// TIA Portal V21 program export: 0 tag tables, 0 data types, 1 data blocks, 40 code blocks (in call order from the OBs), 24 instance data blocks

DATA_BLOCK "Global_Limits_Interlocks"   // DB58
{ S7_Optimized_Access := 'TRUE' }
// stored: MemoryReserve 100
   VAR
      ExternalLevel_Interlock : Real := 2900.0;
      InternalLevel_Interlock : Real := 2700.0;
   END_VAR
BEGIN
END_DATA_BLOCK

ORGANIZATION_BLOCK "Main_1"   // OB1, LAD, ProgramCycle
TITLE = "Main Program Sweep (Cycle)"
{ S7_Optimized_Access := 'TRUE' }
// stored: SetENOAutomatically false
   VAR_INPUT
      Initial_Call : Bool;   // Initial call of this OB
      Remanence : Bool;   // =True, if remanent data are available
   END_VAR
BEGIN
END_ORGANIZATION_BLOCK

ORGANIZATION_BLOCK "Cyclic interrupt"   // OB30, FBD, CyclicInterrupt
{ S7_Optimized_Access := 'TRUE' }
// stored: SetENOAutomatically false
   VAR_INPUT
      Initial_Call : Bool;   // Initial call of this OB
      Event_Count : Int;   // Events discarded
   END_VAR
BEGIN

REGION Network 1: Service
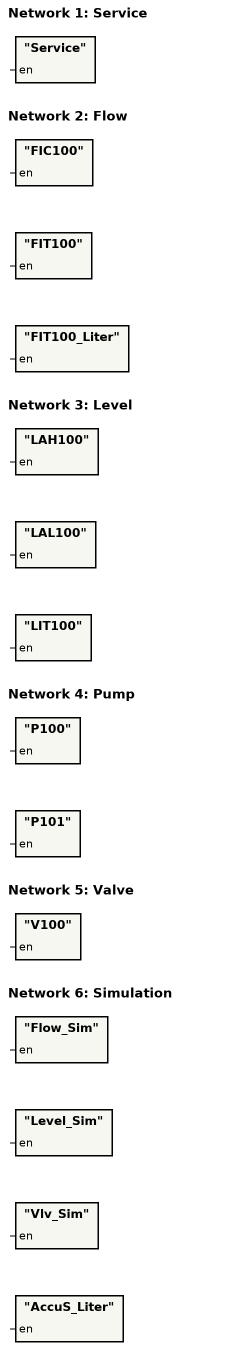
   "Service"();
END_REGION

REGION Network 2: Flow
   "FIC100"();
   "FIT100"();
   "FIT100_Liter"();
END_REGION

REGION Network 3: Level
   "LAH100"();
   "LAL100"();
   "LIT100"();
END_REGION

REGION Network 4: Pump
   "P100"();
   "P101"();
END_REGION

REGION Network 5: Valve
   "V100"();
END_REGION

REGION Network 6: Simulation
   "Flow_Sim"();
   "Level_Sim"();
   "Vlv_Sim"();
   "AccuS_Liter"();
END_REGION
END_ORGANIZATION_BLOCK

FUNCTION "Service" : Void   // FC11, FBD
TITLE = Service
{ S7_Optimized_Access := 'TRUE' }
AUTHOR : Siemens AG
FAMILY : ServiceControl
VERSION : 1.0
// stored: SetENOAutomatically false
   VAR_TEMP
      ProcedureDone : Bool;
      UnholdingDone : Bool;
      StartingState : Bool;
      CompletingState : Bool;
      PausingState : Bool;
      HoldingState : Bool;
      AbortingState : Bool;
      StoppingState : Bool;
      State : "Service_States";
   END_VAR
   VAR_TEMP   // added for the SCL form of the ladder/FBD networks
      _w1 : Bool;
      _w2 : Bool;
      _w3 : Bool;
      _w4 : Bool;
   END_VAR
BEGIN

REGION Network 1: Parameters and values
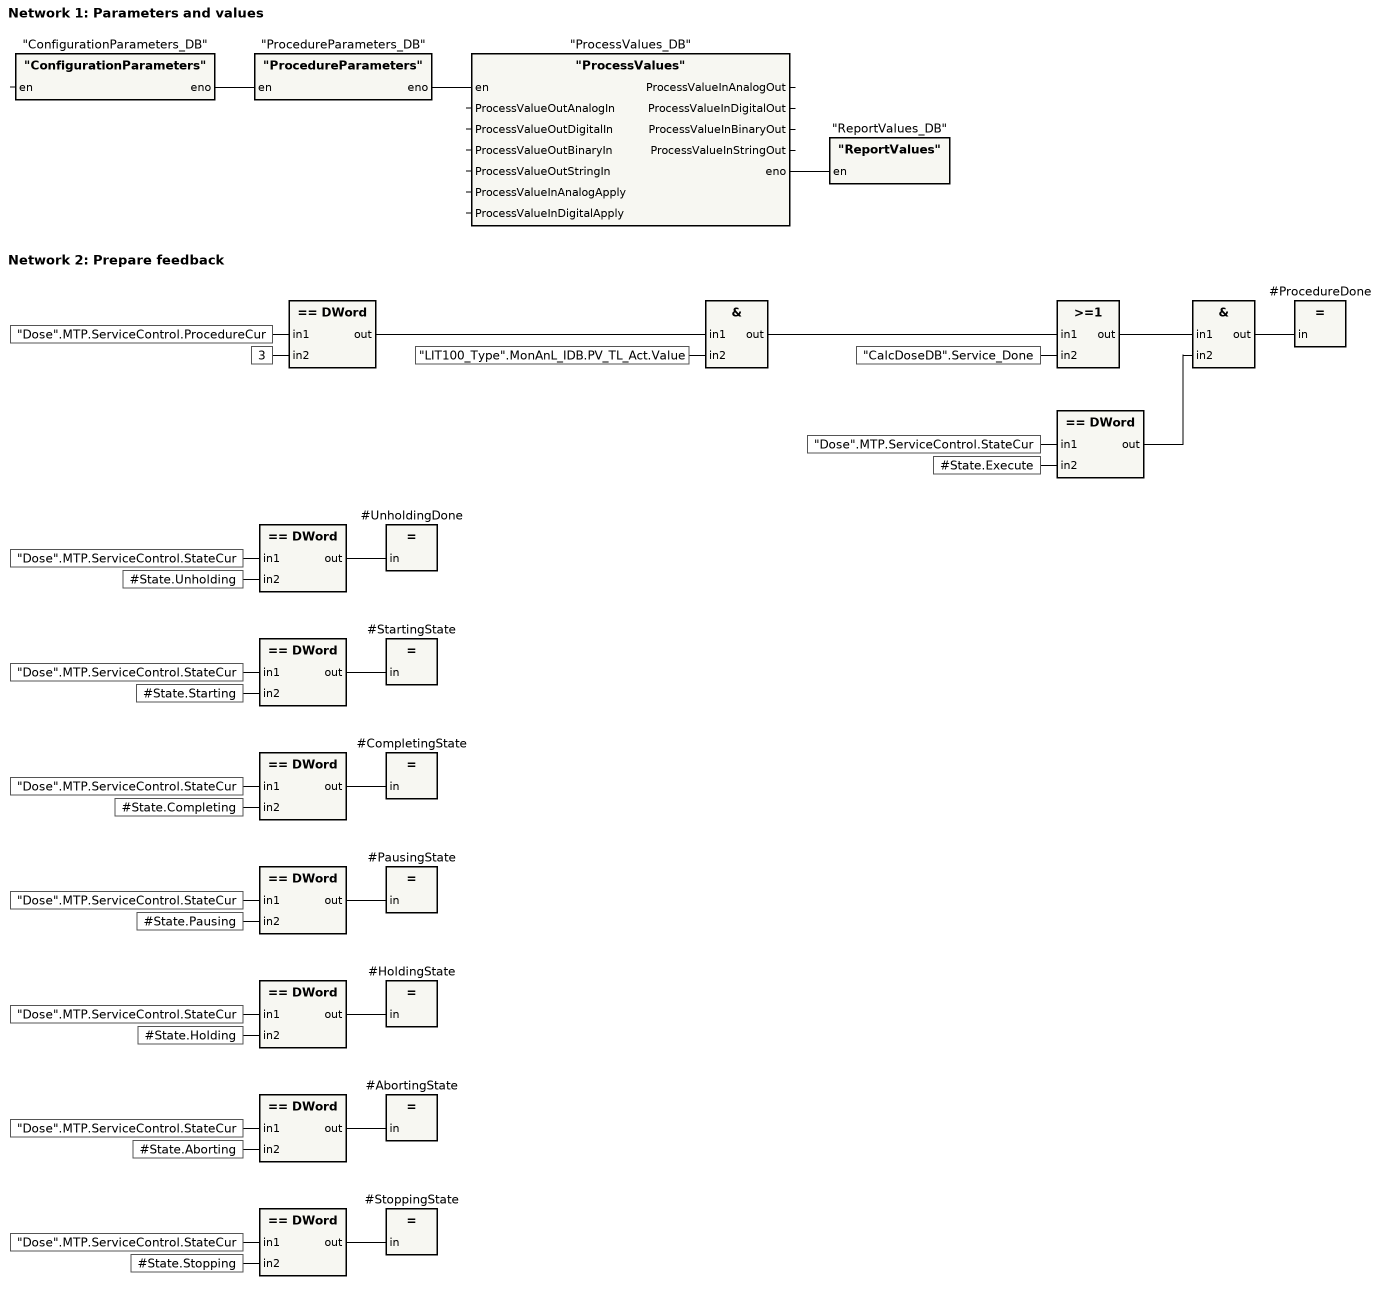
   "ConfigurationParameters_DB"(ENO => #_w1);   // "ConfigurationParameters"
   "ProcedureParameters_DB"(EN := #_w1, ENO => #_w2);   // "ProcedureParameters"
   "ProcessValues_DB"(EN := #_w2, ENO => #_w3);   // "ProcessValues"
   IF #_w3 THEN
       "ReportValues_DB"();   // "ReportValues"
   END_IF;
END_REGION

REGION Network 2: Prepare feedback
   #ProcedureDone := ((("Dose".MTP.ServiceControl.ProcedureCur = 3) AND "LIT100_Type".MonAnL_IDB.PV_TL_Act.Value) OR "CalcDoseDB".Service_Done) AND ("Dose".MTP.ServiceControl.StateCur = #State.Execute);
   #UnholdingDone := "Dose".MTP.ServiceControl.StateCur = #State.Unholding;
   #StartingState := "Dose".MTP.ServiceControl.StateCur = #State.Starting;
   #CompletingState := "Dose".MTP.ServiceControl.StateCur = #State.Completing;
   #PausingState := "Dose".MTP.ServiceControl.StateCur = #State.Pausing;
   #HoldingState := "Dose".MTP.ServiceControl.StateCur = #State.Holding;
   #AbortingState := "Dose".MTP.ServiceControl.StateCur = #State.Aborting;
   #StoppingState := "Dose".MTP.ServiceControl.StateCur = #State.Stopping;
END_REGION

REGION Network 3: Cm P100 feedback
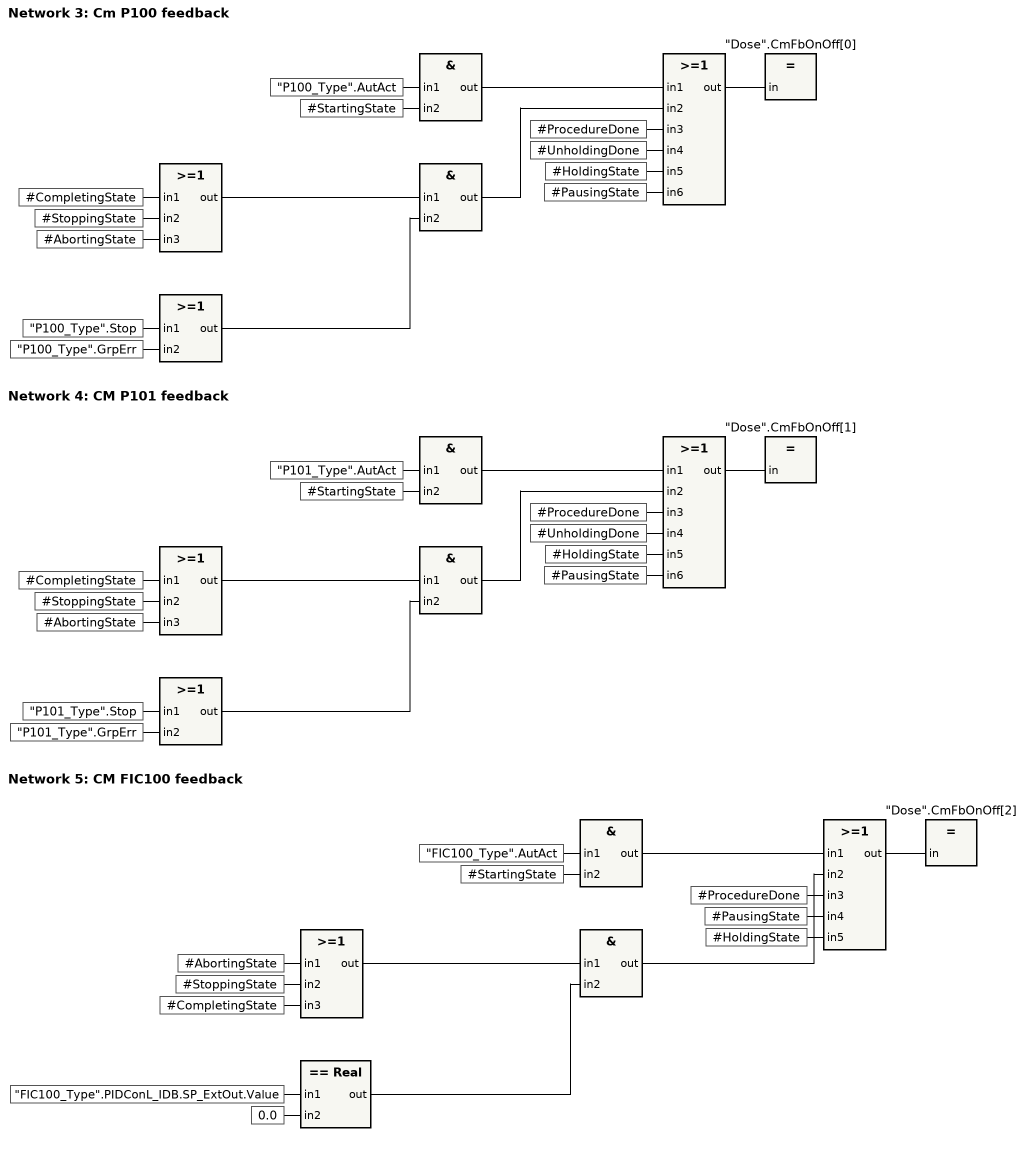
   "Dose".CmFbOnOff[0] := ("P100_Type".AutAct AND #StartingState) OR ((#CompletingState OR #StoppingState OR #AbortingState) AND ("P100_Type".Stop OR "P100_Type".GrpErr)) OR #ProcedureDone OR #UnholdingDone OR #HoldingState OR #PausingState;
END_REGION

REGION Network 4: CM P101 feedback
   "Dose".CmFbOnOff[1] := ("P101_Type".AutAct AND #StartingState) OR ((#CompletingState OR #StoppingState OR #AbortingState) AND ("P101_Type".Stop OR "P101_Type".GrpErr)) OR #ProcedureDone OR #UnholdingDone OR #HoldingState OR #PausingState;
END_REGION

REGION Network 5: CM FIC100 feedback
   "Dose".CmFbOnOff[2] := ("FIC100_Type".AutAct AND #StartingState) OR ((#AbortingState OR #StoppingState OR #CompletingState) AND ("FIC100_Type".PIDConL_IDB.SP_ExtOut.Value = 0.0)) OR #ProcedureDone OR #PausingState OR #HoldingState;
END_REGION

REGION Network 6: CM V100 feedback
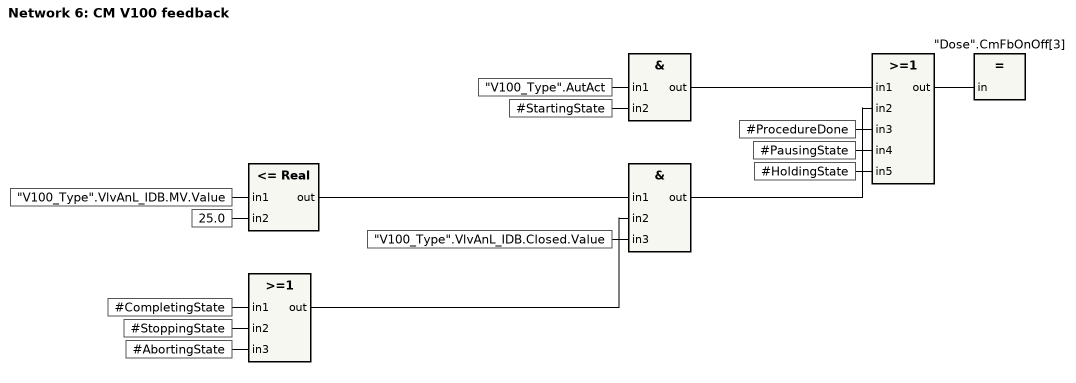
   "Dose".CmFbOnOff[3] := ("V100_Type".AutAct AND #StartingState) OR (("V100_Type".VlvAnL_IDB.MV.Value <= 25.0) AND (#CompletingState OR #StoppingState OR #AbortingState) AND "V100_Type".VlvAnL_IDB.Closed.Value) OR #ProcedureDone OR #PausingState OR #HoldingState;
END_REGION

REGION Network 7: Service
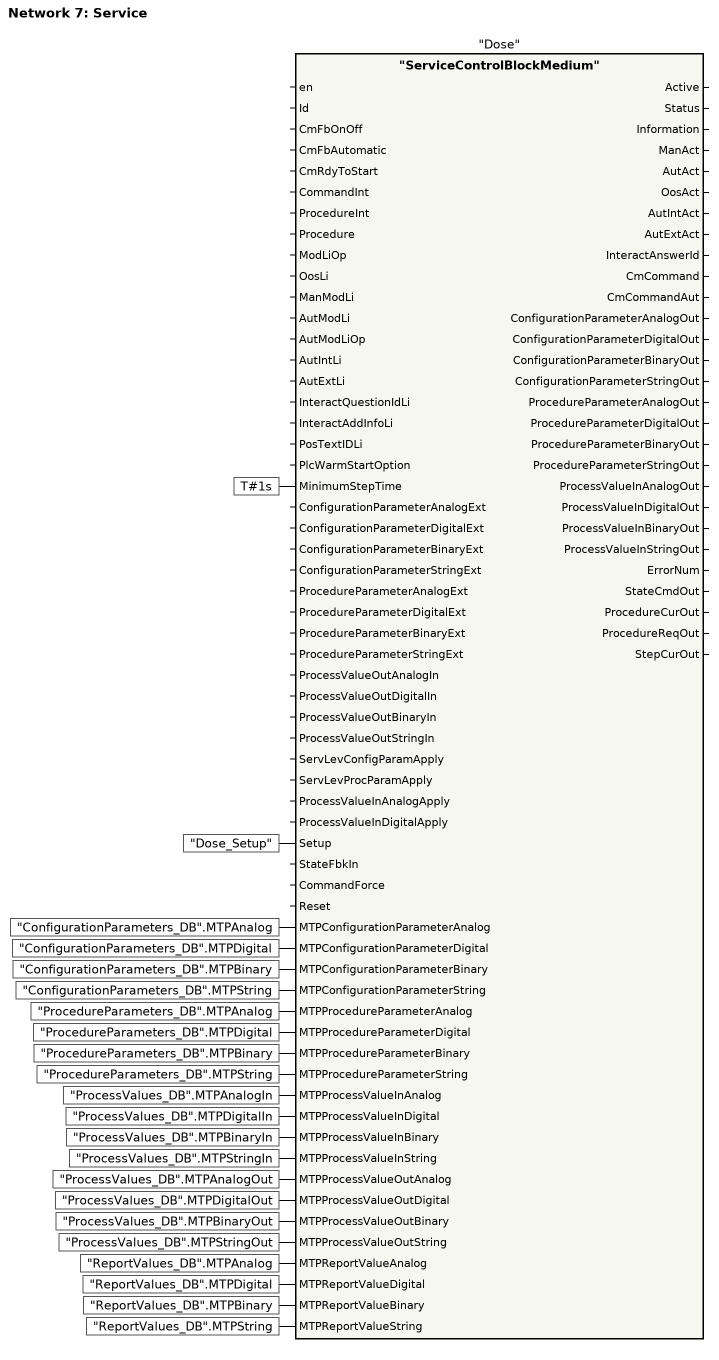
   "Dose"(MinimumStepTime := T#1s,   // "ServiceControlBlockMedium"
          Setup := "Dose_Setup",
          MTPConfigurationParameterAnalog := "ConfigurationParameters_DB".MTPAnalog,
          MTPConfigurationParameterDigital := "ConfigurationParameters_DB".MTPDigital,
          MTPConfigurationParameterBinary := "ConfigurationParameters_DB".MTPBinary,
          MTPConfigurationParameterString := "ConfigurationParameters_DB".MTPString,
          MTPProcedureParameterAnalog := "ProcedureParameters_DB".MTPAnalog,
          MTPProcedureParameterDigital := "ProcedureParameters_DB".MTPDigital,
          MTPProcedureParameterBinary := "ProcedureParameters_DB".MTPBinary,
          MTPProcedureParameterString := "ProcedureParameters_DB".MTPString,
          MTPProcessValueInAnalog := "ProcessValues_DB".MTPAnalogIn,
          MTPProcessValueInDigital := "ProcessValues_DB".MTPDigitalIn,
          MTPProcessValueInBinary := "ProcessValues_DB".MTPBinaryIn,
          MTPProcessValueInString := "ProcessValues_DB".MTPStringIn,
          MTPProcessValueOutAnalog := "ProcessValues_DB".MTPAnalogOut,
          MTPProcessValueOutDigital := "ProcessValues_DB".MTPDigitalOut,
          MTPProcessValueOutBinary := "ProcessValues_DB".MTPBinaryOut,
          MTPProcessValueOutString := "ProcessValues_DB".MTPStringOut,
          MTPReportValueAnalog := "ReportValues_DB".MTPAnalog,
          MTPReportValueDigital := "ReportValues_DB".MTPDigital,
          MTPReportValueBinary := "ReportValues_DB".MTPBinary,
          MTPReportValueString := "ReportValues_DB".MTPString);
END_REGION

REGION Network 8: Service HMI
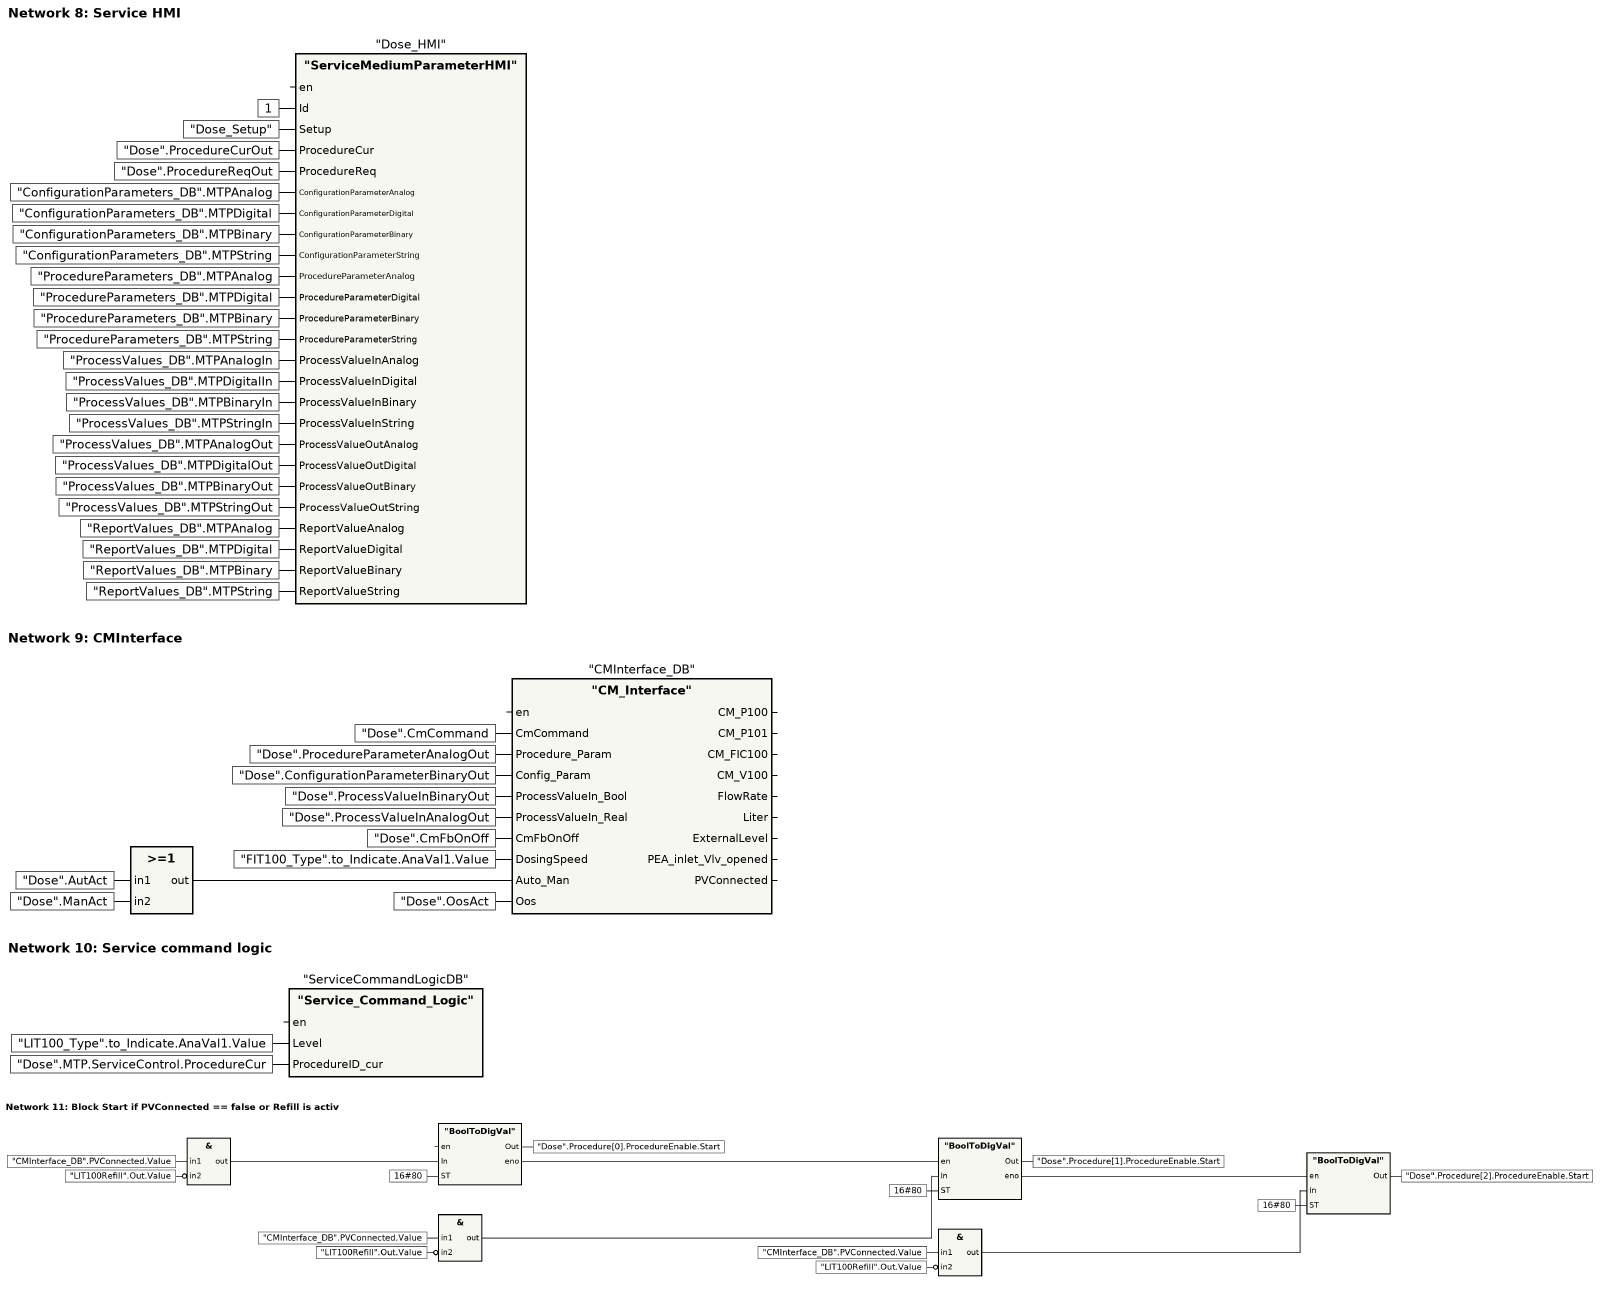
   "Dose_HMI"(Id := 1,   // "ServiceMediumParameterHMI"
              Setup := "Dose_Setup",
              ProcedureCur := "Dose".ProcedureCurOut,
              ProcedureReq := "Dose".ProcedureReqOut,
              ConfigurationParameterAnalog := "ConfigurationParameters_DB".MTPAnalog,
              ConfigurationParameterDigital := "ConfigurationParameters_DB".MTPDigital,
              ConfigurationParameterBinary := "ConfigurationParameters_DB".MTPBinary,
              ConfigurationParameterString := "ConfigurationParameters_DB".MTPString,
              ProcedureParameterAnalog := "ProcedureParameters_DB".MTPAnalog,
              ProcedureParameterDigital := "ProcedureParameters_DB".MTPDigital,
              ProcedureParameterBinary := "ProcedureParameters_DB".MTPBinary,
              ProcedureParameterString := "ProcedureParameters_DB".MTPString,
              ProcessValueInAnalog := "ProcessValues_DB".MTPAnalogIn,
              ProcessValueInDigital := "ProcessValues_DB".MTPDigitalIn,
              ProcessValueInBinary := "ProcessValues_DB".MTPBinaryIn,
              ProcessValueInString := "ProcessValues_DB".MTPStringIn,
              ProcessValueOutAnalog := "ProcessValues_DB".MTPAnalogOut,
              ProcessValueOutDigital := "ProcessValues_DB".MTPDigitalOut,
              ProcessValueOutBinary := "ProcessValues_DB".MTPBinaryOut,
              ProcessValueOutString := "ProcessValues_DB".MTPStringOut,
              ReportValueAnalog := "ReportValues_DB".MTPAnalog,
              ReportValueDigital := "ReportValues_DB".MTPDigital,
              ReportValueBinary := "ReportValues_DB".MTPBinary,
              ReportValueString := "ReportValues_DB".MTPString);
END_REGION

REGION Network 9: CMInterface
   "CMInterface_DB"(CmCommand := "Dose".CmCommand,   // "CM_Interface"
                    Procedure_Param := "Dose".ProcedureParameterAnalogOut,
                    Config_Param := "Dose".ConfigurationParameterBinaryOut,
                    ProcessValueIn_Bool := "Dose".ProcessValueInBinaryOut,
                    ProcessValueIn_Real := "Dose".ProcessValueInAnalogOut,
                    CmFbOnOff := "Dose".CmFbOnOff,
                    DosingSpeed := "FIT100_Type".to_Indicate.AnaVal1.Value,
                    Auto_Man := "Dose".AutAct OR "Dose".ManAct,
                    Oos := "Dose".OosAct);
END_REGION

REGION Network 10: Service command logic
   "ServiceCommandLogicDB"(Level := "LIT100_Type".to_Indicate.AnaVal1.Value,   // "Service_Command_Logic"
                           ProcedureID_cur := "Dose".MTP.ServiceControl.ProcedureCur);
END_REGION

REGION Network 11: Block Start if PVConnected == false or Refill is activ
   "BoolToDigVal"(In := "CMInterface_DB".PVConnected.Value AND NOT "LIT100Refill".Out.Value,
                  ST := 16#80,
                  Out => "Dose".Procedure[0].ProcedureEnable.Start,
                  ENO => #_w1);
   "BoolToDigVal"(EN := #_w1,
                  In := "CMInterface_DB".PVConnected.Value AND NOT "LIT100Refill".Out.Value,
                  ST := 16#80,
                  Out => "Dose".Procedure[1].ProcedureEnable.Start,
                  ENO => #_w2);
   IF #_w2 THEN
       "BoolToDigVal"(In := "CMInterface_DB".PVConnected.Value AND NOT "LIT100Refill".Out.Value,
                      ST := 16#80,
                      Out => "Dose".Procedure[2].ProcedureEnable.Start);
   END_IF;
END_REGION

REGION Network 12: Block Resume and Unholding if refill is activ
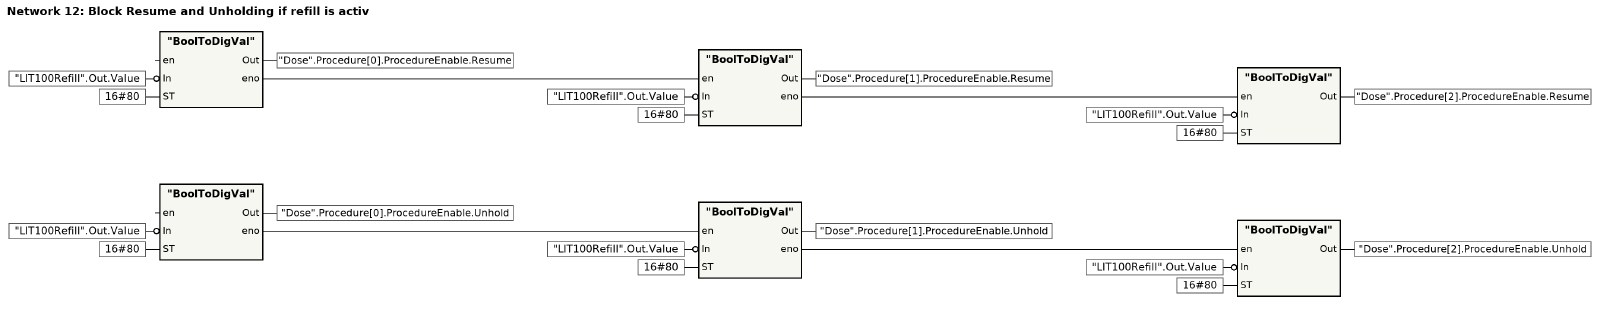
   "BoolToDigVal"(In := NOT "LIT100Refill".Out.Value,
                  ST := 16#80,
                  Out => "Dose".Procedure[0].ProcedureEnable.Resume,
                  ENO => #_w1);
   "BoolToDigVal"(EN := #_w1,
                  In := NOT "LIT100Refill".Out.Value,
                  ST := 16#80,
                  Out => "Dose".Procedure[1].ProcedureEnable.Resume,
                  ENO => #_w2);
   IF #_w2 THEN
       "BoolToDigVal"(In := NOT "LIT100Refill".Out.Value,
                      ST := 16#80,
                      Out => "Dose".Procedure[2].ProcedureEnable.Resume);
   END_IF;
   "BoolToDigVal"(In := NOT "LIT100Refill".Out.Value,
                  ST := 16#80,
                  Out => "Dose".Procedure[0].ProcedureEnable.Unhold,
                  ENO => #_w3);
   "BoolToDigVal"(EN := #_w3,
                  In := NOT "LIT100Refill".Out.Value,
                  ST := 16#80,
                  Out => "Dose".Procedure[1].ProcedureEnable.Unhold,
                  ENO => #_w4);
   IF #_w4 THEN
       "BoolToDigVal"(In := NOT "LIT100Refill".Out.Value,
                      ST := 16#80,
                      Out => "Dose".Procedure[2].ProcedureEnable.Unhold);
   END_IF;
END_REGION

REGION Network 13: Position Text
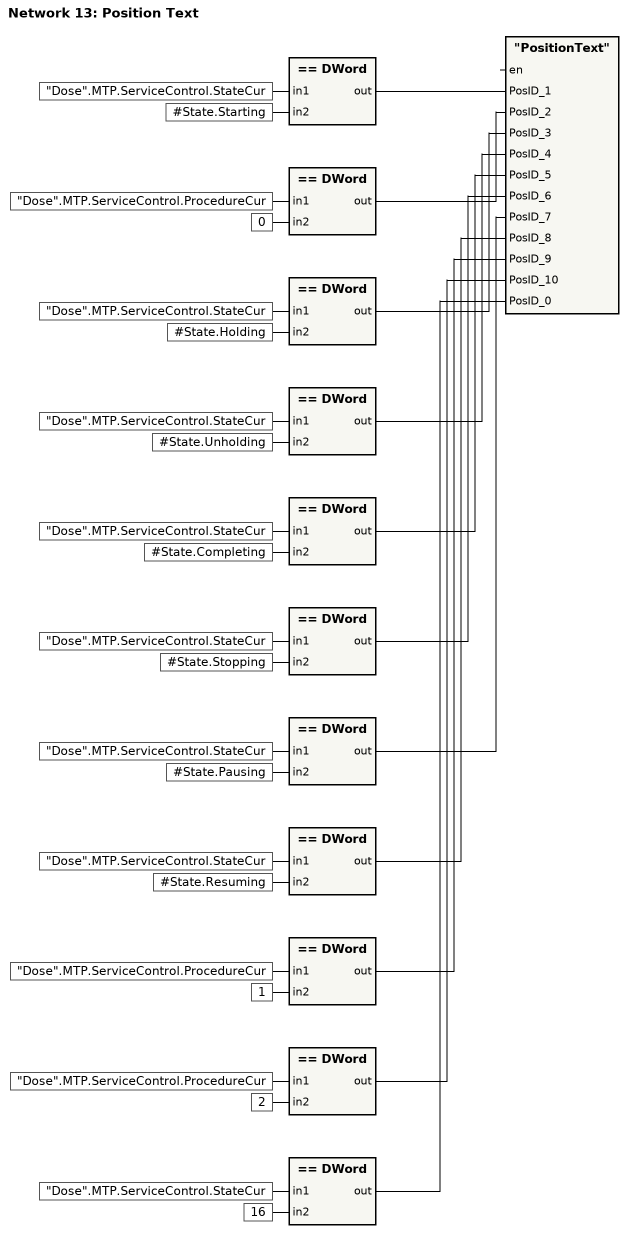
   "PositionText"(PosID_1 := "Dose".MTP.ServiceControl.StateCur = #State.Starting,
                  PosID_2 := "Dose".MTP.ServiceControl.ProcedureCur = 0,
                  PosID_3 := "Dose".MTP.ServiceControl.StateCur = #State.Holding,
                  PosID_4 := "Dose".MTP.ServiceControl.StateCur = #State.Unholding,
                  PosID_5 := "Dose".MTP.ServiceControl.StateCur = #State.Completing,
                  PosID_6 := "Dose".MTP.ServiceControl.StateCur = #State.Stopping,
                  PosID_7 := "Dose".MTP.ServiceControl.StateCur = #State.Pausing,
                  PosID_8 := "Dose".MTP.ServiceControl.StateCur = #State.Resuming,
                  PosID_9 := "Dose".MTP.ServiceControl.ProcedureCur = 1,
                  PosID_10 := "Dose".MTP.ServiceControl.ProcedureCur = 2,
                  PosID_0 := "Dose".MTP.ServiceControl.StateCur = 16);
END_REGION

REGION Network 14: Report values
END_REGION
END_FUNCTION

FUNCTION_BLOCK "ConfigurationParameters"   // FB1710, SCL
TITLE = ConfigurationParameters
{ S7_Optimized_Access := 'TRUE' }
AUTHOR : Siemens AG
FAMILY : ServiceControl
VERSION : 1.0
// Providing of the MTP-Interface and the number of parameters of each configuration parameter type
// stored: MemoryReserve 100, SetENOAutomatically false
   VAR
      MTPAnalog { S7_SetPoint := 'True'} : Array[0..#NUMBER_PARAMETERS_ANALOG] of "UDT_MTP_AnaServParam";
      MTPDigital { S7_SetPoint := 'True'} : Array[0..#NUMBER_PARAMETERS_DIGITAL] of "UDT_MTP_DIntServParam";
      MTPBinary { S7_SetPoint := 'True'} : Array[0..#NUMBER_PARAMETERS_BINARY] of "UDT_MTP_BinServParam";
      MTPString { S7_SetPoint := 'True'} : Array[0..#NUMBER_PARAMETERS_STRING] of "UDT_MTP_StringServParam";
   END_VAR
   VAR CONSTANT
      NUMBER_PARAMETERS_ANALOG : Int := 0;
      NUMBER_PARAMETERS_DIGITAL : Int := 0;
      NUMBER_PARAMETERS_BINARY : Int := 1;
      NUMBER_PARAMETERS_STRING : Int := 0;
   END_VAR
BEGIN
   REGION Block Info Header
     //===============================================================================
     // Siemens AG / (c)Copyright 2021
     //-------------------------------------------------------------------------------
     // Title:            ConfigurationParameters
     // Comment/Function: Providing of the MTP-Interface and the number of parameters of each configuration parameter type
     // Library/Family:   ServiceControl
     // Author:           Siemens AG
     // Tested with:      S7-PLCSIM Advanced 4.0
     // Engineering:      TIA Portal V17
     // Restrictions:     MTP
     // Requirements:     PLC (S7-1200 / S7-1500)
     //-------------------------------------------------------------------------------
     // Change log table:
     // Version  | Date       | Expert in charge        | Changes applied
     //----------|------------|-------------------------|-----------------------------
     // 01.00.00 | 02.09.2021 | Michael Schlosser       | First released version
     // 01.00.01 | 07.09.2021 | Michael Schlosser       | Change: Interface of FB28 ConfigurationParameterAnalog
     // 01.00.02 | 08.09.2021 | Michael Schlosser       | Change: Interface of FB18, FB33, FB24
     // 01.00.03 | 09.09.2021 | Michael Schlosser       | Change: For-loops only until #NUMBER_PARAMETERS_YXZ - 1
     // 01.00.04 | 15.09.2021 | Michael Schlosser       | Change: ApplyEn default values = true (e.g. parLevAnalogApplyEn[0])
     // 01.00.05 | 16.09.2021 | Michael Schlosser       | Change: ApplyEn & ApplyInt as part of UDT_Service_ParameterApply (e.g. #ParLevAnalogApply[0].En)
     // 01.00.06 | 18.10.2021 | Michael Schlosser       | change: call of FBs for parameters now in ServiceControlBlock-FBs to allow several services per PLC
     //===============================================================================
   END_REGION Block Info Header

   REGION Description
     // ConfigurationParameters provides the MTP-Interface and the number of parameters of each configuration parameter type
   END_REGION Description
END_FUNCTION_BLOCK

FUNCTION_BLOCK "ProcedureParameters"   // FB1715, SCL
TITLE = ProcedureParameters
{ S7_Optimized_Access := 'TRUE' }
AUTHOR : Siemens AG
FAMILY : ServiceControl
VERSION : 1.0
// Providing of the MTP-Interface and the number of parameters of each procedure parameter type
// stored: MemoryReserve 100, SetENOAutomatically false
   VAR
      MTPAnalog { S7_SetPoint := 'True'} : Array[0..#NUMBER_PARAMETERS_ANALOG] of "UDT_MTP_AnaServParam";
      MTPDigital { S7_SetPoint := 'True'} : Array[0..#NUMBER_PARAMETERS_DIGITAL] of "UDT_MTP_DIntServParam";
      MTPBinary { S7_SetPoint := 'True'} : Array[0..#NUMBER_PARAMETERS_BINARY] of "UDT_MTP_BinServParam";
      MTPString { S7_SetPoint := 'True'} : Array[0..#NUMBER_PARAMETERS_STRING] of "UDT_MTP_StringServParam";
   END_VAR
   VAR CONSTANT
      NUMBER_PARAMETERS_ANALOG : Int := 2;
      NUMBER_PARAMETERS_DIGITAL : Int := 0;
      NUMBER_PARAMETERS_BINARY : Int := 0;
      NUMBER_PARAMETERS_STRING : Int := 0;
   END_VAR
BEGIN
   REGION Block Info Header
     //===============================================================================
     // Siemens AG / (c)Copyright 2021
     //-------------------------------------------------------------------------------
     // Title:            ProcedureParameters
     // Comment/Function: Providing of the MTP-Interface and the number of parameters of each procedure parameter type
     // Library/Family:   ServiceControl
     // Author:           Siemens AG
     // Tested with:      S7-PLCSIM Advanced 4.0
     // Engineering:      TIA Portal V17
     // Restrictions:     MTP
     // Requirements:     PLC (S7-1200 / S7-1500)
     //-------------------------------------------------------------------------------
     // Change log table:
     // Version  | Date       | Expert in charge        | Changes applied
     //----------|------------|-------------------------|-----------------------------
     // 01.00.00 | 02.09.2021 | Michael Schlosser       | First released version
     // 01.00.01 | 13.09.2021 | Michael Schlosser       | Change: Interface of FB29
     // 01.00.02 | 15.09.2021 | Michael Schlosser       | Change: Interface of FB13, FB19, FB23
     // 01.00.03 | 15.09.2021 | Michael Schlosser       | Change: ApplyEn default values = true (e.g. parLevAnalogApplyEn[0])
     // 01.00.04 | 16.09.2021 | Michael Schlosser       | Change: ApplyEn & ApplyInt as part of UDT_Service_ParameterApply (e.g. #ParLevAnalogApply[0].En)
     // 01.00.05 | 18.10.2021 | Michael Schlosser       | change: call of FBs for parameters now in ServiceControlBlock-FBs to allow several services per PLC
     //===============================================================================
   END_REGION Block Info Header

   REGION Description
     // ProcedureParameters provides the MTP-Interface and the number of parameters of each procedure parameter type
   END_REGION Description
END_FUNCTION_BLOCK

FUNCTION_BLOCK "ProcessValues"   // FB1720, SCL
TITLE = ProcessValues
{ S7_Optimized_Access := 'TRUE' }
AUTHOR : Siemens AG
FAMILY : ServiceControl
VERSION : 1.0
// Handling of ProcessValues
// stored: MemoryReserve 100, SetENOAutomatically false
   VAR_INPUT
      ProcessValueOutAnalogIn { ExternalAccessible := 'False'; ExternalVisible := 'False'; ExternalWritable := 'False'} : Array[0..#NUMBER_PARAMETERS_OUT_ANALOG_NOT_MAPPED] of "UDT_MTP_AnaProcessValueOut";
      ProcessValueOutDigitalIn { ExternalAccessible := 'False'; ExternalVisible := 'False'; ExternalWritable := 'False'} : Array[0..#NUMBER_PARAMETERS_OUT_DIGITAL_NOT_MAPPED] of "UDT_MTP_DIntProcessValueOut";
      ProcessValueOutBinaryIn { ExternalAccessible := 'False'; ExternalVisible := 'False'; ExternalWritable := 'False'} : Array[0..#NUMBER_PARAMETERS_OUT_BINARY_NOT_MAPPED] of "UDT_MTP_BinProcessValueOut";
      ProcessValueOutStringIn { ExternalAccessible := 'False'; ExternalVisible := 'False'; ExternalWritable := 'False'} : Array[0..#NUMBER_PARAMETERS_OUT_STRING_NOT_MAPPED] of "UDT_MTP_StringProcessValueOut";
      ProcessValueInAnalogApply { ExternalAccessible := 'False'; ExternalVisible := 'False'; ExternalWritable := 'False'} : Array[0..#NUMBER_PARAMETERS_IN_ANALOG_NOT_MAPPED] of "UDT_Service_ProcessValueInApply";
      ProcessValueInDigitalApply { ExternalAccessible := 'False'; ExternalVisible := 'False'; ExternalWritable := 'False'} : Array[0..#NUMBER_PARAMETERS_IN_DIGITAL_NOT_MAPPED] of "UDT_Service_ProcessValueInApply";
   END_VAR
   VAR_OUTPUT
      ProcessValueInAnalogOut { ExternalAccessible := 'False'; ExternalVisible := 'False'; ExternalWritable := 'False'} : Array[0..#NUMBER_PARAMETERS_IN_ANALOG_NOT_MAPPED] of "UDT_MTP_AnaProcessValueOut";
      ProcessValueInDigitalOut { ExternalAccessible := 'False'; ExternalVisible := 'False'; ExternalWritable := 'False'} : Array[0..#NUMBER_PARAMETERS_IN_DIGITAL_NOT_MAPPED] of "UDT_MTP_DIntProcessValueOut";
      ProcessValueInBinaryOut { ExternalAccessible := 'False'; ExternalVisible := 'False'; ExternalWritable := 'False'} : Array[0..#NUMBER_PARAMETERS_IN_BINARY_NOT_MAPPED] of "UDT_MTP_BinProcessValueOut";
      ProcessValueInStringOut { ExternalAccessible := 'False'; ExternalVisible := 'False'; ExternalWritable := 'False'} : Array[0..#NUMBER_PARAMETERS_IN_STRING_NOT_MAPPED] of "UDT_MTP_StringProcessValueOut";
   END_VAR
   VAR
      MTPAnalogIn : Array[0..#NUMBER_PARAMETERS_IN_ANALOG_TOTAL] of "UDT_MTP_AnaProcessValueIn";
      MTPDigitalIn : Array[0..#NUMBER_PARAMETERS_IN_DIGITAL_TOTAL] of "UDT_MTP_DIntProcessValueIn";
      MTPBinaryIn : Array[0..#NUMBER_PARAMETERS_IN_BINARY_TOTAL] of "UDT_MTP_BinProcessValueIn";
      MTPStringIn : Array[0..#NUMBER_PARAMETERS_IN_STRING_TOTAL] of "UDT_MTP_StringProcessValueIn";
      AnalogIn { ExternalAccessible := 'False'; ExternalVisible := 'False'; ExternalWritable := 'False'; S7_SetPoint := 'True'} : Array[0..#NUMBER_PARAMETERS_IN_ANALOG_NOT_MAPPED] of "ProcessValueInAnalog";
      DigitalIn { ExternalAccessible := 'False'; ExternalVisible := 'False'; ExternalWritable := 'False'; S7_SetPoint := 'True'} : Array[0..#NUMBER_PARAMETERS_IN_DIGITAL_NOT_MAPPED] of "ProcessValueInDigital";
      BinaryIn { ExternalAccessible := 'False'; ExternalVisible := 'False'; ExternalWritable := 'False'; S7_SetPoint := 'True'} : Array[0..#NUMBER_PARAMETERS_IN_BINARY_NOT_MAPPED] of "ProcessValueInBinary";
      StringIn { ExternalAccessible := 'False'; ExternalVisible := 'False'; ExternalWritable := 'False'; S7_SetPoint := 'True'} : Array[0..#NUMBER_PARAMETERS_IN_STRING_NOT_MAPPED] of "ProcessValueInString";
      MTPAnalogOut : Array[0..#NUMBER_PARAMETERS_OUT_ANALOG_TOTAL] of "UDT_MTP_AnaProcessValueOut";
      MTPDigitalOut : Array[0..#NUMBER_PARAMETERS_OUT_DIGITAL_TOTAL] of "UDT_MTP_DIntProcessValueOut";
      MTPBinaryOut : Array[0..#NUMBER_PARAMETERS_OUT_BINARY_TOTAL] of "UDT_MTP_BinProcessValueOut";
      MTPStringOut : Array[0..#NUMBER_PARAMETERS_OUT_STRING_TOTAL] of "UDT_MTP_StringProcessValueOut";
      AnalogOut { ExternalAccessible := 'False'; ExternalVisible := 'False'; ExternalWritable := 'False'; S7_SetPoint := 'True'} : Array[0..#NUMBER_PARAMETERS_OUT_ANALOG_NOT_MAPPED] of "ProcessValueOutAnalog";
      DigitalOut { ExternalAccessible := 'False'; ExternalVisible := 'False'; ExternalWritable := 'False'; S7_SetPoint := 'True'} : Array[0..#NUMBER_PARAMETERS_OUT_DIGITAL_NOT_MAPPED] of "ProcessValueOutDigital";
      BinaryOut { ExternalAccessible := 'False'; ExternalVisible := 'False'; ExternalWritable := 'False'; S7_SetPoint := 'True'} : Array[0..#NUMBER_PARAMETERS_OUT_BINARY_NOT_MAPPED] of "ProcessValueOutBinary";
      StringOut { ExternalAccessible := 'False'; ExternalVisible := 'False'; ExternalWritable := 'False'; S7_SetPoint := 'True'} : Array[0..#NUMBER_PARAMETERS_OUT_STRING_NOT_MAPPED] of "ProcessValueOutString";
   END_VAR
   VAR_TEMP
      i : Int;
      tempUpperLimit : Int;   // Upper limit for FOR - loop
      tempModuloNumber : Int;   // Number for modulo calculation
      tempIndexExt : Int;   // Index for external interface of not mapped process values
      tempTVO : Bool;   // Transfer value only from Ext to MTP (instead of whole UDT)
   END_VAR
   VAR CONSTANT
      NUMBER_PARAMETERS_IN_ANALOG_TOTAL : Int := 1;
      NUMBER_PARAMETERS_IN_DIGITAL_TOTAL : Int := 0;
      NUMBER_PARAMETERS_IN_BINARY_TOTAL : Int := 1;
      NUMBER_PARAMETERS_IN_STRING_TOTAL : Int := 0;
      NUMBER_PARAMETERS_OUT_ANALOG_TOTAL : Int := 1;
      NUMBER_PARAMETERS_OUT_DIGITAL_TOTAL : Int := 0;
      NUMBER_PARAMETERS_OUT_BINARY_TOTAL : Int := 0;
      NUMBER_PARAMETERS_OUT_STRING_TOTAL : Int := 0;
      NUMBER_PARAMETERS_IN_ANALOG_NOT_MAPPED : Int;   // Not mapped to a service
      NUMBER_PARAMETERS_IN_DIGITAL_NOT_MAPPED : Int;   // Not mapped to a service
      NUMBER_PARAMETERS_IN_BINARY_NOT_MAPPED : Int;   // Not mapped to a service
      NUMBER_PARAMETERS_IN_STRING_NOT_MAPPED : Int;   // Not mapped to a service
      NUMBER_PARAMETERS_OUT_ANALOG_NOT_MAPPED : Int;   // Not mapped to a service
      NUMBER_PARAMETERS_OUT_DIGITAL_NOT_MAPPED : Int;   // Not mapped to a service
      NUMBER_PARAMETERS_OUT_BINARY_NOT_MAPPED : Int;   // Not mapped to a service
      NUMBER_PARAMETERS_OUT_STRING_NOT_MAPPED : Int;   // Not mapped to a service
      NUMBER_PARAMETERS_IN_MIN : Int;
      NUMBER_PARAMETERS_OUT_MIN : Int;
   END_VAR
BEGIN
   REGION Block Info Header
     //===============================================================================
     // Siemens AG / (c)Copyright 2021
     //-------------------------------------------------------------------------------
     // Title:            ProcessValues
     // Comment/Function: Handling of ProcessValues
     // Library/Family:   ServiceControl
     // Author:           Siemens AG
     // Tested with:      S7-PLCSIM Advanced 4.0
     // Engineering:      TIA Portal V17
     // Restrictions:     MTP
     // Requirements:     PLC (S7-1200 / S7-1500)
     //-------------------------------------------------------------------------------
     // Change log table:
     // Version  | Date       | Expert in charge        | Changes applied
     //----------|------------|-------------------------|-----------------------------
     // 01.00.00 | 29.07.2021 | Michael Schlosser       | First released version
     // 01.00.01 | 20.09.2021 | Michael Schlosser       | change: comment in region "Description"; new comments of for-loops
     // 01.00.02 | 19.10.2021 | Markus Krause           | change: New Outputs for PV Inputs without Service
     // 01.00.03 | 21.10.2021 | Markus Krause           | change: New concept for Standalone mode of the Process Values Inputs / Outputs
     // 01.00.04 | 22.10.2021 | Markus Krause           | change: Bugfix for Standalone mode of the Process Values Inputs / Outputs
     // 01.00.05 | 22.10.2021 | Markus Krause           | change: Bugfix for Standalone mode of the Process Values Inputs / Outputs
     // 01.00.06 | 22.10.2021 | Markus Krause           | change: ApplyEn changed from Bool to UDT_Service_ProcessValueInApply
     // 01.00.07 | 25.10.2021 | Michael Schlosser       | change: process out values are now connected via InOut interface "Ext" to process value out FBs
     // 01.00.08 | 26.10.2021 | Michael Schlosser       | change: differentiation between "mapped" and "not mapped" for process values out
     // 01.00.09 | 27.10.2021 | Michael Schlosser       | change: process in values are now connected via InOut interface "Ext" to process value in FBs; differentiation between "mapped" and "not mapped" for process values in
     // 01.00.10 | 28.10.2021 | Michael Schlosser       | rename: interface "isMapped" to "TVO" (transfer value only) for process values out
     // 01.00.11 | 22.11.2021 | Michael Schlosser       | change: extend comment in region "Description"
     //===============================================================================
   END_REGION Block Info Header

   REGION Description
     // ProcessValues provides the MTP-Interface and the number of values of each type of process in/out value
     // and calls the FB for each analog, digital, binary and string process in/out value which is not mapped to any service
   END_REGION Description

   REGION BLOCK INITIALIZATION
     #tempTVO := false;  // Transfer whole UDT from Ext to MTP for not mapped (to a service) process values out
   END_REGION BLOCK INITIALIZATION

   REGION BEHAVIOR LOGIC

     // Call of process value FB for each not mapped analog in value
     #tempUpperLimit := #NUMBER_PARAMETERS_IN_ANALOG_TOTAL - 1 + #NUMBER_PARAMETERS_IN_MIN;
     #tempModuloNumber := #NUMBER_PARAMETERS_IN_ANALOG_TOTAL;  // without this trick, the compiler throws error division by zero 
     FOR #i := #NUMBER_PARAMETERS_IN_MIN TO #tempUpperLimit DO
       IF (#i > #tempUpperLimit - #NUMBER_PARAMETERS_IN_ANALOG_NOT_MAPPED) AND (#tempModuloNumber > 0) AND (#tempModuloNumber >= #NUMBER_PARAMETERS_IN_ANALOG_NOT_MAPPED) THEN
         // Number_Mapped + Number_not_Mapped = Number_Total
         // Call FB only in case that the values of the constants are consistent and that no division by zero is possible
         #tempIndexExt := ((#i + #NUMBER_PARAMETERS_IN_ANALOG_NOT_MAPPED) MOD #tempModuloNumber) + #NUMBER_PARAMETERS_IN_MIN;
         // Not-mapped (to a service) process values in are located at upper MTP-indices and must be mapped to their external output area
         #AnalogIn[#tempIndexExt](Apply := #ProcessValueInAnalogApply[#tempIndexExt],
                                  MTP   := #MTPAnalogIn[#i],
                                  Ext   := #ProcessValueInAnalogOut[#tempIndexExt]);
       END_IF;
     END_FOR;

     // Call of process value FB for each not mapped digital in value
     #tempUpperLimit := #NUMBER_PARAMETERS_IN_DIGITAL_TOTAL - 1 + #NUMBER_PARAMETERS_IN_MIN;
     #tempModuloNumber := #NUMBER_PARAMETERS_IN_DIGITAL_TOTAL;  // without this trick, the compiler throws error division by zero 
     FOR #i := #NUMBER_PARAMETERS_IN_MIN TO #tempUpperLimit DO
       IF (#i > #tempUpperLimit - #NUMBER_PARAMETERS_IN_DIGITAL_NOT_MAPPED) AND (#tempModuloNumber > 0) AND (#tempModuloNumber >= #NUMBER_PARAMETERS_IN_DIGITAL_NOT_MAPPED) THEN
         // Number_Mapped + Number_not_Mapped = Number_Total
         // Call FB only in case that the values of the constants are consistent and that no division by zero is possible
         #tempIndexExt := ((#i + #NUMBER_PARAMETERS_IN_DIGITAL_NOT_MAPPED) MOD #tempModuloNumber) + #NUMBER_PARAMETERS_IN_MIN;
         // Not-mapped (to a service) process values in are located at upper MTP-indices and must be mapped to their external output area
         #DigitalIn[#tempIndexExt](Apply := #ProcessValueInDigitalApply[#tempIndexExt],
                                   MTP   := #MTPDigitalIn[#i],
                                   Ext   := #ProcessValueInDigitalOut[#tempIndexExt]);
       END_IF;
     END_FOR;

     // Call of process value FB for each not mapped binary in value
     #tempUpperLimit := #NUMBER_PARAMETERS_IN_BINARY_TOTAL - 1 + #NUMBER_PARAMETERS_IN_MIN;
     #tempModuloNumber := #NUMBER_PARAMETERS_IN_BINARY_TOTAL;  // without this trick, the compiler throws error division by zero 
     FOR #i := #NUMBER_PARAMETERS_IN_MIN TO #tempUpperLimit DO
       IF (#i > #tempUpperLimit - #NUMBER_PARAMETERS_IN_BINARY_NOT_MAPPED) AND (#tempModuloNumber > 0) AND (#tempModuloNumber >= #NUMBER_PARAMETERS_IN_BINARY_NOT_MAPPED) THEN
         // Number_Mapped + Number_not_Mapped = Number_Total
         // Call FB only in case that the values of the constants are consistent and that no division by zero is possible
         #tempIndexExt := ((#i + #NUMBER_PARAMETERS_IN_BINARY_NOT_MAPPED) MOD #tempModuloNumber) + #NUMBER_PARAMETERS_IN_MIN;
         // Not-mapped (to a service) process values in are located at upper MTP-indices and must be mapped to their external output area
         #BinaryIn[#tempIndexExt](MTP := #MTPBinaryIn[#i],
                                  Ext := #ProcessValueInBinaryOut[#tempIndexExt]);
       END_IF;
     END_FOR;

     // Call of process value FB for each not mapped string in value
     #tempUpperLimit := #NUMBER_PARAMETERS_IN_STRING_TOTAL - 1 + #NUMBER_PARAMETERS_IN_MIN;
     #tempModuloNumber := #NUMBER_PARAMETERS_IN_STRING_TOTAL;  // without this trick, the compiler throws error division by zero 
     FOR #i := #NUMBER_PARAMETERS_IN_MIN TO #tempUpperLimit DO
       IF (#i > #tempUpperLimit - #NUMBER_PARAMETERS_IN_STRING_NOT_MAPPED) AND (#tempModuloNumber > 0) AND (#tempModuloNumber >= #NUMBER_PARAMETERS_IN_STRING_NOT_MAPPED) THEN
         // Number_Mapped + Number_not_Mapped = Number_Total
         // Call FB only in case that the values of the constants are consistent and that no division by zero is possible
         #tempIndexExt := ((#i + #NUMBER_PARAMETERS_IN_STRING_NOT_MAPPED) MOD #tempModuloNumber) + #NUMBER_PARAMETERS_IN_MIN;
         // Not-mapped (to a service) process values in are located at upper MTP-indices and must be mapped to their external output area
         #StringIn[#tempIndexExt](MTP := #MTPStringIn[#i],
                                  Ext := #ProcessValueInStringOut[#tempIndexExt]);
       END_IF;
     END_FOR;



     // Call of process value FB for each not mapped analog out value
     #tempUpperLimit := #NUMBER_PARAMETERS_OUT_ANALOG_TOTAL - 1 + #NUMBER_PARAMETERS_OUT_MIN;
     #tempModuloNumber := #NUMBER_PARAMETERS_OUT_ANALOG_TOTAL;  // without this trick, the compiler throws error division by zero 
     FOR #i := #NUMBER_PARAMETERS_OUT_MIN TO #tempUpperLimit DO
       IF (#i > #tempUpperLimit - #NUMBER_PARAMETERS_OUT_ANALOG_NOT_MAPPED) AND (#tempModuloNumber > 0) AND (#tempModuloNumber >= #NUMBER_PARAMETERS_OUT_ANALOG_NOT_MAPPED) THEN
         // Number_Mapped + Number_not_Mapped = Number_Total
         // Call FB only in case that the values of the constants are consistent and that no division by zero is possible
         #tempIndexExt := ((#i + #NUMBER_PARAMETERS_OUT_ANALOG_NOT_MAPPED) MOD #tempModuloNumber) + #NUMBER_PARAMETERS_OUT_MIN;
         // Not-mapped (to a service) process values out are located at upper MTP-indices and must be mapped to their external input area
         #AnalogOut[#tempIndexExt](TVO := #tempTVO,
                                   Ext := #ProcessValueOutAnalogIn[#tempIndexExt],
                                   MTP := #MTPAnalogOut[#i]);
       END_IF;
     END_FOR;

     // Call of process value FB for each not mapped digital out value
     #tempUpperLimit := #NUMBER_PARAMETERS_OUT_DIGITAL_TOTAL - 1 + #NUMBER_PARAMETERS_OUT_MIN;
     #tempModuloNumber := #NUMBER_PARAMETERS_OUT_DIGITAL_TOTAL;  // without this trick, the compiler throws error division by zero 
     FOR #i := #NUMBER_PARAMETERS_OUT_MIN TO #tempUpperLimit DO
       IF (#i > #tempUpperLimit - #NUMBER_PARAMETERS_OUT_DIGITAL_NOT_MAPPED) AND (#tempModuloNumber > 0) AND (#tempModuloNumber >= #NUMBER_PARAMETERS_OUT_DIGITAL_NOT_MAPPED) THEN
         // Number_Mapped + Number_not_Mapped = Number_Total
         // Call FB only in case that the values of the constants are consistent and that no division by zero is possible
         #tempIndexExt := ((#i + #NUMBER_PARAMETERS_OUT_DIGITAL_NOT_MAPPED) MOD #tempModuloNumber) + #NUMBER_PARAMETERS_OUT_MIN;
         // Not-mapped (to a service) process values out are located at upper MTP-indices and must be mapped to their external input area
         #DigitalOut[#tempIndexExt](TVO := #tempTVO,
                                    Ext := #ProcessValueOutDigitalIn[#tempIndexExt],
                                    MTP := #MTPDigitalOut[#i]);
       END_IF;
     END_FOR;

     // Call of process value FB for each not mapped binary out value
     #tempUpperLimit := #NUMBER_PARAMETERS_OUT_BINARY_TOTAL - 1 + #NUMBER_PARAMETERS_OUT_MIN;
     #tempModuloNumber := #NUMBER_PARAMETERS_OUT_BINARY_TOTAL;  // without this trick, the compiler throws error division by zero 
     FOR #i := #NUMBER_PARAMETERS_OUT_MIN TO #tempUpperLimit DO
       IF (#i > #tempUpperLimit - #NUMBER_PARAMETERS_OUT_BINARY_NOT_MAPPED) AND (#tempModuloNumber > 0) AND (#tempModuloNumber >= #NUMBER_PARAMETERS_OUT_BINARY_NOT_MAPPED) THEN
         // Number_Mapped + Number_not_Mapped = Number_Total
         // Call FB only in case that the values of the constants are consistent and that no division by zero is possible
         #tempIndexExt := ((#i + #NUMBER_PARAMETERS_OUT_BINARY_NOT_MAPPED) MOD #tempModuloNumber) + #NUMBER_PARAMETERS_OUT_MIN;
         // Not-mapped (to a service) process values out are located at upper MTP-indices and must be mapped to their external input area
         #BinaryOut[#tempIndexExt](TVO := #tempTVO,
                                   Ext := #ProcessValueOutBinaryIn[#tempIndexExt],
                                   MTP := #MTPBinaryOut[#i]);
       END_IF;
     END_FOR;

     // Call of process value FB for each not mapped string out value
     #tempUpperLimit := #NUMBER_PARAMETERS_OUT_STRING_TOTAL - 1 + #NUMBER_PARAMETERS_OUT_MIN;
     #tempModuloNumber := #NUMBER_PARAMETERS_OUT_STRING_TOTAL;  // without this trick, the compiler throws error division by zero 
     FOR #i := #NUMBER_PARAMETERS_OUT_MIN TO #tempUpperLimit DO
       IF (#i > #tempUpperLimit - #NUMBER_PARAMETERS_OUT_STRING_NOT_MAPPED) AND (#tempModuloNumber > 0) AND (#tempModuloNumber >= #NUMBER_PARAMETERS_OUT_STRING_NOT_MAPPED) THEN
         // Number_Mapped + Number_not_Mapped = Number_Total
         // Call FB only in case that the values of the constants are consistent and that no division by zero is possible
         #tempIndexExt := ((#i + #NUMBER_PARAMETERS_OUT_STRING_NOT_MAPPED) MOD #tempModuloNumber) + #NUMBER_PARAMETERS_OUT_MIN;
         // Not-mapped (to a service) process values out are located at upper MTP-indices and must be mapped to their external input area
         #StringOut[#tempIndexExt](TVO := #tempTVO,
                                   Ext := #ProcessValueOutStringIn[#tempIndexExt],
                                   MTP := #MTPStringOut[#i]);
       END_IF;
     END_FOR;

   END_REGION BEHAVIOR LOGIC
END_FUNCTION_BLOCK

FUNCTION_BLOCK "ReportValues"   // FB1730, SCL
TITLE = ReportValues
{ S7_Optimized_Access := 'TRUE' }
AUTHOR : Siemens AG
FAMILY : ServiceControl
VERSION : 1.0
// Handling of ReportValues
// stored: MemoryReserve 100, SetENOAutomatically false
   VAR
      MTPAnalog { S7_SetPoint := 'True'} : Array[0..#NUMBER_PARAMETERS_ANALOG] of "UDT_MTP_AnaReportValue";
      MTPDigital { S7_SetPoint := 'True'} : Array[0..#NUMBER_PARAMETERS_DIGITAL] of "UDT_MTP_DIntReportValue";
      MTPBinary { S7_SetPoint := 'True'} : Array[0..#NUMBER_PARAMETERS_BINARY] of "UDT_MTP_BinReportValue";
      MTPString { S7_SetPoint := 'True'} : Array[0..#NUMBER_PARAMETERS_STRING] of "UDT_MTP_StringReportValue";
   END_VAR
   VAR CONSTANT
      NUMBER_PARAMETERS_ANALOG : Int := 1;
      NUMBER_PARAMETERS_DIGITAL : Int := 0;
      NUMBER_PARAMETERS_BINARY : Int := 0;
      NUMBER_PARAMETERS_STRING : Int := 0;
   END_VAR
BEGIN
   REGION Block Info Header
     //===============================================================================
     // Siemens AG / (c)Copyright 2021
     //-------------------------------------------------------------------------------
     // Title:            ReportValues
     // Comment/Function: Handling of ReportValues
     // Library/Family:   ServiceControl
     // Author:           Siemens AG
     // Tested with:      S7-PLCSIM Advanced 4.0
     // Engineering:      TIA Portal V17
     // Restrictions:     MTP
     // Requirements:     PLC (S7-1200 / S7-1500)
     //-------------------------------------------------------------------------------
     // Change log table:
     // Version  | Date       | Expert in charge        | Changes applied
     //----------|------------|-------------------------|-----------------------------
     // 01.00.00 | 29.07.2021 | Michael Schlosser       | First released version
     // 01.00.01 | 21.09.2021 | Michael Schlosser       | change: comment in region "Description"; new comments of for-loops
     // 01.00.02 | 21.10.2021 | Michael Schlosser       | change: call of FBs for report values now in ServiceControlBlock-FBs to allow several services per PLC
     //===============================================================================
   END_REGION Block Info Header

   REGION Description
     // ReportValues provides the MTP-Interface and the number of values of each type of report value
   END_REGION Description
END_FUNCTION_BLOCK

FUNCTION_BLOCK "ServiceMediumParameterHMI"   // FB1754, SCL
TITLE = ServiceMediumParameterHMI
{ S7_Optimized_Access := 'TRUE' }
AUTHOR : Siemens AG
FAMILY : ServiceControl
VERSION : 4.0
// { "TagName" : "" , "TagDescription" : "" }
// stored: MemoryReserve 100, SetENOAutomatically false
   VAR_INPUT
      Id { ExternalAccessible := 'False'; ExternalVisible := 'False'; ExternalWritable := 'False'} : USInt;   // Service parameter ID
      Setup { ExternalAccessible := 'False'; ExternalVisible := 'False'; ExternalWritable := 'False'} : DB_ANY;   // Setup DB used for the service
      ProcedureCur { ExternalAccessible := 'False'; ExternalVisible := 'False'; ExternalWritable := 'False'} : DWord;   // Current Procedure Number
      ProcedureReq { ExternalAccessible := 'False'; ExternalVisible := 'False'; ExternalWritable := 'False'} : DWord;   // Required Procedure Numbar
   END_VAR
   VAR_IN_OUT
      ConfigurationParameterAnalog : Array[*] of "UDT_MTP_AnaServParam";   // Analog configuration parameter
      ConfigurationParameterDigital : Array[*] of "UDT_MTP_DIntServParam";   // Digital configuration parameter
      ConfigurationParameterBinary : Array[*] of "UDT_MTP_BinServParam";   // Binary configuration parameter
      ConfigurationParameterString : Array[*] of "UDT_MTP_StringServParam";   // String configuration parameter
      ProcedureParameterAnalog : Array[*] of "UDT_MTP_AnaServParam";   // Analog configuration parameter / Analog procedure parameter
      ProcedureParameterDigital : Array[*] of "UDT_MTP_DIntServParam";   // Digital configuration parameter / Digital procedure parameter
      ProcedureParameterBinary : Array[*] of "UDT_MTP_BinServParam";   // Binary configuration parameter / Binary procedure parameter
      ProcedureParameterString : Array[*] of "UDT_MTP_StringServParam";   // String configuration parameter / String procedure parameter
      ProcessValueInAnalog : Array[*] of "UDT_MTP_AnaProcessValueIn";   // Analog process value in
      ProcessValueInDigital : Array[*] of "UDT_MTP_DIntProcessValueIn";   // Digital process value in
      ProcessValueInBinary : Array[*] of "UDT_MTP_BinProcessValueIn";   // Binary process value in
      ProcessValueInString : Array[*] of "UDT_MTP_StringProcessValueIn";   // String process value in
      ProcessValueOutAnalog : Array[*] of "UDT_MTP_AnaProcessValueOut";   // Analog process value out
      ProcessValueOutDigital : Array[*] of "UDT_MTP_DIntProcessValueOut";   // Digital process value out
      ProcessValueOutBinary : Array[*] of "UDT_MTP_BinProcessValueOut";   // Binary process value out
      ProcessValueOutString : Array[*] of "UDT_MTP_StringProcessValueOut";   // String process value out
      ReportValueAnalog : Array[*] of "UDT_MTP_AnaReportValue";   // Analog report value
      ReportValueDigital : Array[*] of "UDT_MTP_DIntReportValue";   // Digital report value
      ReportValueBinary : Array[*] of "UDT_MTP_BinReportValue";   // Binary report value
      ReportValueString : Array[*] of "UDT_MTP_StringReportValue";   // String report value
   END_VAR
   VAR
      statTotalConfigParameters { ExternalAccessible := 'False'; ExternalVisible := 'False'; ExternalWritable := 'False'} : Int;   // Total used configuration parameter
      statTotalProcedureParameters { ExternalAccessible := 'False'; ExternalVisible := 'False'; ExternalWritable := 'False'} : Int;   // Total used procedure parameter
      statTotalProcessInValues { ExternalAccessible := 'False'; ExternalVisible := 'False'; ExternalWritable := 'False'} : Int;   // Total used process in values
      statTotalProcessOutValues { ExternalAccessible := 'False'; ExternalVisible := 'False'; ExternalWritable := 'False'} : Int;   // Total used process Out values
      statTotalReportValues { ExternalAccessible := 'False'; ExternalVisible := 'False'; ExternalWritable := 'False'} : Int;   // Total used Report values
      StatConfigAnalog { ExternalAccessible := 'False'; ExternalVisible := 'False'; ExternalWritable := 'False'} : Array[0..#MAPPED_CONFIG_ANALOG] of "UDT_Service_AnaServParam";   // Writable Config analog parameters
      StatConfigDigital { ExternalAccessible := 'False'; ExternalVisible := 'False'; ExternalWritable := 'False'} : Array[0..#MAPPED_CONFIG_DIGITAL] of "UDT_Service_DintServParam";   // Writable Config digital parameters
      StatConfigBinary { ExternalAccessible := 'False'; ExternalVisible := 'False'; ExternalWritable := 'False'} : Array[0..#MAPPED_CONFIG_BINARY] of "UDT_Service_BinServParam";   // Writable Config binary parameters
      StatConfigString { ExternalAccessible := 'False'; ExternalVisible := 'False'; ExternalWritable := 'False'} : Array[0..#MAPPED_CONFIG_STRING] of "UDT_Service_StringServParam";   // Writable Config string parameters
      StatProcedureAnalog { ExternalAccessible := 'False'; ExternalVisible := 'False'; ExternalWritable := 'False'} : Array[0..#MAPPED_PROCEDURE_ANALOG] of "UDT_Service_AnaServParam";   // Writable Config analog parameters
      StatProcedureDigital { ExternalAccessible := 'False'; ExternalVisible := 'False'; ExternalWritable := 'False'} : Array[0..#MAPPED_PROCEDURE_DIGITAL] of "UDT_Service_DintServParam";   // Writable Config digital parameters
      StatProcedureBinary { ExternalAccessible := 'False'; ExternalVisible := 'False'; ExternalWritable := 'False'} : Array[0..#MAPPED_PROCEDURE_BINARY] of "UDT_Service_BinServParam";   // Writable Config binary parameters
      StatProcedureString { ExternalAccessible := 'False'; ExternalVisible := 'False'; ExternalWritable := 'False'} : Array[0..#MAPPED_PROCEDURE_STRING] of "UDT_Service_StringServParam";   // Writable Config string parameters
      stat16ProceReqIndex { ExternalAccessible := 'False'; ExternalVisible := 'False'; ExternalWritable := 'False'} : Int;   // Requested/Prepared procedure index number
      stat16ProceCurIndex { ExternalAccessible := 'False'; ExternalVisible := 'False'; ExternalWritable := 'False'} : Int;   // current/Running procedure index number
      stat16ProcParaStartIndex { ExternalAccessible := 'False'; ExternalVisible := 'False'; ExternalWritable := 'False'} : Int;   // Procedure parameter start index value
      stat16ProcParaEndIndex { ExternalAccessible := 'False'; ExternalVisible := 'False'; ExternalWritable := 'False'} : Int;   // Procedure parameter end index value
      stat32PrecedureProcessOutMap { ExternalAccessible := 'False'; ExternalVisible := 'False'; ExternalWritable := 'False'} : DWord;   // Procedure assignment information for ProcessOut values
      stat32PrecedureProcessInMap { ExternalAccessible := 'False'; ExternalVisible := 'False'; ExternalWritable := 'False'} : DWord;   // Procedure assignment information for ProcessIn values
      stat32PrecedureReportMap { ExternalAccessible := 'False'; ExternalVisible := 'False'; ExternalWritable := 'False'} : DWord;   // Procedure assignment information for Report values
      ConfigParaType : "UDT_Service_ConfigParaIndexType";   // Index information for the configuration parameter
      ProcedureParaType : "UDT_Service_ProceParaValueIndexType";   // Index information for the procedure parameter
      ProcessInValueType : "UDT_Service_ProceParaValueIndexType";   // Index information for the process in values
      ProcessOutValueType : "UDT_Service_ProceParaValueIndexType";   // Index information for the process out values
      ReportValueType : "UDT_Service_ProceParaValueIndexType";   // Index information for the report values
      ConfigAna : Array[0..#MAPPED_CONFIG_ANALOG] of "UDT_MTP_AnaServParam";   // Configuration analog parameter
      ConfigDint : Array[0..#MAPPED_CONFIG_DIGITAL] of "UDT_MTP_DIntServParam";   // Configuration digital parameter
      ConfigBin : Array[0..#MAPPED_CONFIG_BINARY] of "UDT_MTP_BinServParam";   // Configuration binary parameter
      ConfigString : Array[0..#MAPPED_CONFIG_STRING] of "UDT_MTP_StringServParam";   // Configuration string parameter
      ProcedureAna : Array[0..#MAPPED_PROCEDURE_ANALOG] of "UDT_MTP_AnaServParam";   // Procedure analog parameter
      ProcedureDint : Array[0..#MAPPED_PROCEDURE_DIGITAL] of "UDT_MTP_DIntServParam";   // Procedure digital parameter
      ProcedureBin : Array[0..#MAPPED_PROCEDURE_BINARY] of "UDT_MTP_BinServParam";   // Procedure binary parameter
      ProcedureString : Array[0..#MAPPED_PROCEDURE_STRING] of "UDT_MTP_StringServParam";   // Procedure string parameter
      ProcessInAna : Array[0..#MAPPED_PROCESS_IN_ANALOG] of "UDT_MTP_AnaProcessValueIn";   // Process In analog values
      ProcessInDint : Array[0..#MAPPED_PROCESS_IN_DIGITAL] of "UDT_MTP_DIntProcessValueIn";   // Process In digital values
      ProcessInBin : Array[0..#MAPPED_PROCESS_IN_BINARY] of "UDT_MTP_BinProcessValueIn";   // Process In binary values
      ProcessInString : Array[0..#MAPPED_PROCESS_IN_STRING] of "UDT_MTP_StringProcessValueIn";   // Process In string values
      ProcessOutAna : Array[0..#MAPPED_PROCESS_OUT_ANALOG] of "UDT_MTP_AnaProcessValueOut";   // Process Out analog values
      ProcessOutDint : Array[0..#MAPPED_PROCESS_OUT_DIGITAL] of "UDT_MTP_DIntProcessValueOut";   // Process Out digital values
      ProcessOutBin : Array[0..#MAPPED_PROCESS_OUT_BINARY] of "UDT_MTP_BinProcessValueOut";   // Process Out binary values
      ProcessOutString : Array[0..#MAPPED_PROCESS_OUT_STRING] of "UDT_MTP_StringProcessValueOut";   // Process Out string values
      ReportAna : Array[0..#MAPPED_REPORT_ANALOG] of "UDT_MTP_AnaReportValue";   // Report analog values
      ReportDint : Array[0..#MAPPED_REPORT_DIGITAL] of "UDT_MTP_DIntReportValue";   // Report digital values
      ReportBin : Array[0..#MAPPED_REPORT_BINARY] of "UDT_MTP_BinReportValue";   // Report binary values
      ReportString : Array[0..#MAPPED_REPORT_STRING] of "UDT_MTP_StringReportValue";   // Report string values
      statInternalCurProcParameter { ExternalAccessible := 'False'; ExternalVisible := 'False'; ExternalWritable := 'False'} : Array[#PROCEDURE_PARAMETER_MIN..#PROCEDURE_PARAMETER_MAX] of "UDT_Service_Parameter";   // Internal Procedure Parameter
      statLasProcedureCur { ExternalAccessible := 'False'; ExternalVisible := 'False'; ExternalWritable := 'False'} : DWord;   // Last current procedure
      statLasProcedureReq { ExternalAccessible := 'False'; ExternalVisible := 'False'; ExternalWritable := 'False'} : DWord;   // Last Prepared procedure
      statLastReqProcedSelected { ExternalAccessible := 'False'; ExternalVisible := 'False'; ExternalWritable := 'False'} : Bool;   // Last Prepared procedure
      StatLastProceselReport { ExternalAccessible := 'False'; ExternalVisible := 'False'; ExternalWritable := 'False'} : Bool;   // Last procedure page selection in Report values FP
      StatLastProceselProcessOut { ExternalAccessible := 'False'; ExternalVisible := 'False'; ExternalWritable := 'False'} : Bool;   // Last procedure page selection in ProcessOut values FP
      StatLastProceselProcessIn { ExternalAccessible := 'False'; ExternalVisible := 'False'; ExternalWritable := 'False'} : Bool;   // Last procedure page selection in ProcessIn values FP
   END_VAR
   VAR_TEMP
      temp32TempDword1 : DWord;   // Dummy for work
      temp16IndexOfDefinition : Int;   // Index of Definition array / Internal counter variable
      temp16ParameterCMAddress : Int;   // Control module address of parameter
      temp16ParameterType : Int;   // Type of Parameter
      temp16IndexMTP : Int;   // Index of MTP array / Index fo value
      temp16IndexIO : Int;   // Index of IO array / Index fo value
      tempUsed : Array[#NUMBER_OF_CONTROLMODULES_IN_DW_MIN..#NUMBER_OF_CONTROLMODULES_IN_DW] of DWord;   // Array for input value used
      temp16TempInt1 : Int;   // Dummy for work
      temp16TempInt2 : Int;   // Dummy for work
      temp16i : Int;   // Internal counter variable
      temp16Index : Int;   // Index of value / Index fo value
      tempVariant : Variant;   // Internal work variable of type Variant
      temp16ReturnValue : Int;   // Internal work variable for Return Value
      tempSetup : "UDT_Service_ControlBlockMedium";   // Content of DB "ServiceControlBlockMediumSetup"
      tempProcStartIndex : Int;   // Procedure start index
      tempProcEndIndex : Int;   // Procedure end index
      temp16InitIndex : Int;   // Variable is used to initialize the Digital & String para index
      tempProcStartingStartIndex : Int;   // Procedure start index for Starting state
      tempProcStartingEndIndex : Int;   // Procedure end index for Starting state
      tempProcRunningStartIndex : Int;   // Procedure start index for Running state
      tempProcRunningEndIndex : Int;   // Procedure end index for Running state
      tempProcHoldingStartIndex : Int;   // Procedure start index for Holding state
      tempProcHoldingEndIndex : Int;   // Procedure end index for Holding state
      tempProcUnHoldingStartIndex : Int;   // Procedure start index for UnHolding state
      tempProcUnHoldingEndIndex : Int;   // Procedure end index for UnHolding state
      tempProcUnPausingStartIndex : Int;   // Procedure start index for Pausing state
      tempProcUnPausingEndIndex : Int;   // Procedure end index for Pausing state
      tempProcResumingStartIndex : Int;   // Procedure start index for Resuming state
      tempProcResumingEndIndex : Int;   // Procedure end index for Resuming state
      tempProcCompletingStartIndex : Int;   // Procedure start index for Completing state
      tempProcCompletingEndIndex : Int;   // Procedure end index for Completing state
      tempProcStoppingStartIndex : Int;   // Procedure start index for Stopping state
      tempProcStoppingEndIndex : Int;   // Procedure end index for Stopping state
      tempProcAbortingStartIndex : Int;   // Procedure start index for Aborting state
      tempProcAbortingEndIndex : Int;   // Procedure end index for Aborting state
      tempProcResettingStartIndex : Int;   // Procedure start index for Resetting state
      tempProcResettingEndIndex : Int;   // Procedure end index for Resetting state
      temp16IndexOfDefinitionProcessOut : Int;   // Index of Definition array / Internal counter variable
      temp16IndexOfDefinitionProcessIn : Int;   // Index of Definition array / Internal counter variable
      temp16IndexOfDefinitionReport : Int;   // Index of Definition array / Internal counter variable
      temp16IndexAnalog : Int;   // Pointer for the used analog parameter
      temp16IndexDigital : Int;   // Pointer for the used digital parameter
      temp16IndexBinary : Int;   // Pointer for the used binary parameter
      temp16IndexString : Int;   // Pointer for the used string parameter
      temp16ReturnValueOBNum : Int;   // Internal work variable for Return Value
      tempTopSi : SI_none;   // Start-up information of current OB
      tempStartSi : SI_none;   // Start-up information of last started OB
      temp16ObNo : UInt;   // OB number
      xOB_Start : Bool;   // block is running in start OB
      temp16ReturnStatus : Word;   // Internal work variable for Return Value
      tempDTLCurrentTime : DTL;   // Current time stamp
   END_VAR
   VAR CONSTANT
      CONFIG_PARAMETER_MIN : Int := 0;   // Minimum number of configuration parameters (planned number -1 due to ArrayAddressing)
      CONFIG_PARAMETER_MAX : Int := 31;   // Maximum number of configuration parameters (planned number -1 due to ArrayAddressing)
      CONFIG_PARAMETER_ANALOG_MAX : Int := 31;   // Maximum number of analog configuration parameters (planned number -1 due to ArrayAddressing)
      CONFIG_PARAMETER_DIGITAL_MAX : Int := 7;   // Maximum number of digital configuration parameters (planned number -1 due to ArrayAddressing)
      CONFIG_PARAMETER_BINARY_MAX : Int := 31;   // Maximum number of binary configuration parameters (planned number -1 due to ArrayAddressing)
      CONFIG_PARAMETER_STRING_MAX : Int := 7;   // Maximum number of string configuration parameters (planned number -1 due to ArrayAddressing)
      PROCEDURE_PARAMETER_MIN : Int := 0;   // Minimum number of procedure parameters (planned number -1 due to ArrayAddressing)
      PROCEDURE_PARAMETER_MAX : Int := 31;   // Maximum number of procedure parameters (planned number -1 due to ArrayAddressing)
      PROCEDURE_PARAMETER_ANALOG_MAX : Int := 31;   // Maximum number of analog procedure parameters (planned number -1 due to ArrayAddressing)
      PROCEDURE_PARAMETER_DIGITAL_MAX : Int := 7;   // Maximum number of digital procedure parameters (planned number -1 due to ArrayAddressing)
      PROCEDURE_PARAMETER_BINARY_MAX : Int := 31;   // Maximum number of binary procedure parameters (planned number -1 due to ArrayAddressing)
      PROCEDURE_PARAMETER_STRING_MAX : Int := 7;   // Maximum number of string procedure parameters (planned number -1 due to ArrayAddressing)
      NUMBER_OF_CONTROLMODULES_IN_DW_MIN : Int := 0;   // Number of control modules coded in DWords (planned number -1 due to ArrayAddressing)
      NUMBER_OF_CONTROLMODULES_IN_DW : Int := 0;   // Number of control modules coded in DWords (planned number -1 due to ArrayAddressing)
      NUMBER_OF_CONTROLMODULES_MIN : Int := 0;   // Number of control modules (planned number -1 due to ArrayAddressing)
      NUMBER_OF_CONTROLMODULES : Int := 29;   // Number of control modules (planned number -1 due to ArrayAddressing)
      TYPE_NONE : USInt := 0;   // No parameter
      TYPE_ANALOG : USInt := 1;   // Parameter / value type analog
      TYPE_DIGITAL : USInt := 2;   // Parameter / value type digital
      TYPE_BINARY : USInt := 3;   // Parameter / value type binary
      TYPE_STRING : USInt := 4;   // Parameter type string
      NUMBER_OF_PROCEDURES_MIN : Int := 0;   // Number of operations (planned number -1 due to ArrayAddressing)
      NUMBER_OF_PROCEDURES : Int := 15;   // Number of operations (planned number -1 due to ArrayAddressing)
      PARAMETERINDEX_MIN : Int := 0;   // Minimum number of configuration parameters (planned number -1 due to ArrayAddressing)
      PARAMETERINDEX_MAX : Int := 511;   // Maximum number of configuration parameters (planned number -1 due to ArrayAddressing)
      REPORT_VALUES_MIN : Int := 0;   // Minimum number of report values (planned number -1 due to ArrayAddressing)
      REPORT_VALUES_MAX : Int := 31;   // Maximum number of report values (planned number -1 due to ArrayAddressing)
      REPORT_VALUES_ANALOG_MAX : Int := 31;   // Maximum number of analog report values (planned number -1 due to ArrayAddressing)
      REPORT_VALUES_DIGITAL_MAX : Int := 7;   // Maximum number of digital report values (planned number -1 due to ArrayAddressing)
      REPORT_VALUES_BINARY_MAX : Int := 31;   // Maximum number of binary report values (planned number -1 due to ArrayAddressing)
      REPORT_VALUES_STRING_MAX : Int := 7;   // Maximum number of string report values (planned number -1 due to ArrayAddressing)
      PROCESS_VALUES_IN_MIN : Int := 0;   // Minimum number of process values in (planned number -1 due to ArrayAddressing)
      PROCESS_VALUES_IN_MAX : Int := 31;   // Maximum number of process values in (planned number -1 due to ArrayAddressing)
      PROCESS_VALUES_IN_ANALOG_MAX : Int := 31;   // Maximum number of analog process values in (planned number -1 due to ArrayAddressing)
      PROCESS_VALUES_IN_DIGITAL_MAX : Int := 7;   // Maximum number of digital process values in (planned number -1 due to ArrayAddressing)
      PROCESS_VALUES_IN_BINARY_MAX : Int := 31;   // Maximum number of binary process values in (planned number -1 due to ArrayAddressing)
      PROCESS_VALUES_IN_STRING_MAX : Int := 7;   // Maximum number of string process values in (planned number -1 due to ArrayAddressing)
      PROCESS_VALUES_OUT_MIN : Int := 0;   // Minimum number of process values out (planned number -1 due to ArrayAddressing)
      PROCESS_VALUES_OUT_MAX : Int := 31;   // Maximum number of process values out (planned number -1 due to ArrayAddressing)
      PROCESS_VALUES_OUT_ANALOG_MAX : Int := 31;   // Maximum number of analog process values out (planned number -1 due to ArrayAddressing)
      PROCESS_VALUES_OUT_DIGITAL_MAX : Int := 7;   // Maximum number of digital process values out (planned number -1 due to ArrayAddressing)
      PROCESS_VALUES_OUT_BINARY_MAX : Int := 31;   // Maximum number of binary process values out (planned number -1 due to ArrayAddressing)
      PROCESS_VALUES_OUT_STRING_MAX : Int := 7;   // Maximum number of string process values out (planned number -1 due to ArrayAddressing)
      MAPPED_CONFIG_ANALOG : Int := 0;   // Mapped configuration analog parameter count
      MAPPED_CONFIG_DIGITAL : Int := 0;   // Mapped configuration digital parameter count
      MAPPED_CONFIG_BINARY : Int := 1;   // Mapped configuration binary parameter count
      MAPPED_CONFIG_STRING : Int := 0;   // Mapped configuration string parameter count
      MAPPED_PROCEDURE_ANALOG : Int := 2;   // Mapped procedure analog parameter count
      MAPPED_PROCEDURE_DIGITAL : Int := 0;   // Mapped procedure digital parameter count
      MAPPED_PROCEDURE_BINARY : Int := 0;   // Mapped procedure binary parameter count
      MAPPED_PROCEDURE_STRING : Int := 0;   // Mapped procedure string parameter count
      MAPPED_PROCESS_IN_ANALOG : Int := 1;   // Mapped process In analog values count
      MAPPED_PROCESS_IN_DIGITAL : Int := 0;   // Mapped process In Digital values count
      MAPPED_PROCESS_IN_BINARY : Int := 1;   // Mapped process In Binary values count
      MAPPED_PROCESS_IN_STRING : Int := 0;   // Mapped process In String values count
      MAPPED_PROCESS_OUT_ANALOG : Int := 1;   // Mapped process Out analog values count
      MAPPED_PROCESS_OUT_DIGITAL : Int := 0;   // Mapped process Out digital values count
      MAPPED_PROCESS_OUT_BINARY : Int := 0;   // Mapped process Out binary values count
      MAPPED_PROCESS_OUT_STRING : Int := 0;   // Mapped process Out string values count
      MAPPED_REPORT_ANALOG : Int := 1;   // Mapped report analog values count
      MAPPED_REPORT_DIGITAL : Int := 0;   // Mapped report digital values count
      MAPPED_REPORT_BINARY : Int := 0;   // Mapped report binary values count
      MAPPED_REPORT_STRING : Int := 0;   // Mapped report string values count
   END_VAR
BEGIN
       REGION Copyright, Change Log
   (*-----------------------------------------------------------------------------------------------------------------------------
       SIEMENS AG
       © Copyright 2021. All Rights Reserved.
       ---------------------------------------------------------------------------------------------------------------------------
       Limitation of liability
       This software was developed with largest care. However, the author can not
       guarantee, that the software runs under each version of SIMATIC Manager on
       each computer flawlessly. There is no warranty for the software, to the extent
       permitted by applicable law. The copyright holder provides the software
       "as is" without warranty of any kind, either expressed or implied, including,
       but not limited to, the implied warranties of merchantability and fitness
       for a particular purpose. The entire risk as to the quality and performance of
       the software is with you. Should the software prove defective, you assume the
       cost of all necessary servicing, repair or correction. In no event unless
       required by applicable law will the copyright holder be liable to you for
       damages, including any general, special, incidental or consequential damages
       arising out of the use or inability to use the software (including but not
       limited to loss of data or data being rendered inaccurate or losses sustained
       by you or third parties or a failure of the software to operate with any
       other programs), even if such holder or other party has been advised of the
       possibility of such damages. Permission to use or copy this software for any
       purpose is hereby granted without fee, provided the above notices are retained
       on all copies. Permission to modify the code and to distribute modified code
       is granted, provided the above notices are retained, and a notice that the
       code was modified is included with the above copyright notice.
       ---------------------------------------------------------------------------------------------------------------------------
       Functionality provided by this source (short description):
       Function block to handle the Parameters mapped/used in the project from the engineering tool.
       ---------------------------------------------------------------------------------------------------------------------------
       Status: Preliminary,
       Preliminary (experimental)
       Baselined  
       Released
       ---------------------------------------------------------------------------------------------------------------------------
       File name:              ServiceParameter.SCL
       Function block name:    "ServiceParameterFB"
       System :                SIMATIC S7 CPU (1500)
       ---------------------------------------------------------------------------------------------------------------------------
       Restrictions, known limitations: (e.g. only for certain platforms, ...)
       The provided source code is applicable to the CPUs of the S7 1500 series
       ---------------------------------------------------------------------------------------------------------------------------
       Requirements, prerequisites, external resources used: (e.g. hardware,
       technological package, memory needed, other scripts which are included,
       other objects instantiated, other applications (e.g. MS Excel) assumed, ...)
       TIA Version V19
       ---------------------------------------------------------------------------------------------------------------------------
       Change log table (latest change is at the bottom of the list):
        Version  | Date       | Expert in charge        | Changes applied
       ----------|------------|-------------------------|-----------------------------
        00.00.01 | 06.03.2024 | Kumaraguru M            | first implement  
        00.00.11 | 26.03.2024 | Kumaraguru M            | BugFix - 682100 - SPFL Library: When the user creates a procedure without assigning a step in the transit state, and after downloading the file to PLC, PLC goes into STOP mode.  
        03.00.01 | 07.04.2024 | Kumaraguru M            | Feature -676519: Process In value view for Service Control Block 
        03.00.01 | 07.04.2024 | Kumaraguru M            | Feature -676521: Process Out value View for Service Control Block 
        03.00.01 | 07.04.2024 | Kumaraguru M            | Feature -676524: Report Value View for Service Control Block
       ---------------------------------------------------------------------------------------------------------------------------
        27.04.2024 - Changed the FB from Type to Master Copy for Memory and Power Tag Optimization
        08.05.2024 - Change : Bug 702554: SPFL: Service Control Block: In the runtime, when the user has not selected a procedure, then the ProcessIn, Processout, and Report parameters are listed.
        08.05.2024 - Change : Bug 700381: SPFL: SPFL Library: When the user engineers the “ServiceParameterHMI” block icon, the interface tag names are not in uniform.
        12.05.2024 - Change : Bug 702859: SPFL: Service Control Block: In the configuration windows, the parameter values are continuously updated.
       ---------------------------------------------------------------------------------------------------------------------------
       Note:User should not change or modify the logic and interfaces of the Funtion Block.
       ---------------------------------------------------------------------------------------------------------------------------*)
       END_REGION

       REGION Get start information / time information
           #temp16ReturnValueOBNum := RD_SINFO(TOP_SI => #tempTopSi, START_UP_SI => #tempStartSi);
           #temp16ObNo := #tempTopSi.OB_Nr;
           #xOB_Start := false;
           IF (#temp16ObNo = 100) THEN
               #xOB_Start := true;
           END_IF;
           #temp16ReturnStatus := INT_TO_WORD(RD_SYS_T(#tempDTLCurrentTime));

       END_REGION

       REGION Initialization
           IF (#temp16ObNo = 100) THEN
               //Reset Config para index
               #ConfigParaType.IndexAnalog := 16#0;
               #ConfigParaType.IndexDigital := 16#0;
               #ConfigParaType.IndexBinary := 16#0;
               #ConfigParaType.IndexString := 16#0;
               //Reset Procedure para index
               #ProcedureParaType.IndexAnalog := 16#0;
               #ProcedureParaType.NameIndexAnalog := 16#0;
               #ProcedureParaType.IndexDigital := 16#0;
               #ProcedureParaType.NameIndexDigital := 16#0;
               #ProcedureParaType.IndexBinary := 16#0;
               #ProcedureParaType.NameIndexBinary := 16#0;
               #ProcedureParaType.IndexString := 16#0;
               #ProcedureParaType.NameIndexString := 16#0;
               //Reset ProcessIn Value index
               #ProcessInValueType.IndexAnalog := 16#0;
               #ProcessInValueType.NameIndexAnalog := 16#0;
               #ProcessInValueType.IndexDigital := 16#0;
               #ProcessInValueType.NameIndexDigital := 16#0;
               #ProcessInValueType.IndexBinary := 16#0;
               #ProcessInValueType.NameIndexBinary := 16#0;
               #ProcessInValueType.IndexString := 16#0;
               #ProcessInValueType.NameIndexString := 16#0;
               //Reset ProcessOut Value index
               #ProcessOutValueType.IndexAnalog := 16#0;
               #ProcessOutValueType.NameIndexAnalog := 16#0;
               #ProcessOutValueType.IndexDigital := 16#0;
               #ProcessOutValueType.NameIndexDigital := 16#0;
               #ProcessOutValueType.IndexBinary := 16#0;
               #ProcessOutValueType.NameIndexBinary := 16#0;
               #ProcessOutValueType.IndexString := 16#0;
               #ProcessOutValueType.NameIndexString := 16#0;
               //Reset Report Value index
               #ReportValueType.IndexAnalog := 16#0;
               #ReportValueType.NameIndexAnalog := 16#0;
               #ReportValueType.IndexDigital := 16#0;
               #ReportValueType.NameIndexDigital := 16#0;
               #ReportValueType.IndexBinary := 16#0;
               #ReportValueType.NameIndexBinary := 16#0;
               #ReportValueType.IndexString := 16#0;
               #ReportValueType.NameIndexString := 16#0;

           END_IF;
       END_REGION


       REGION Check DB_ANY of Source
           // Get the Setup DB UDT info from the Setup DB 
           #tempVariant := DB_ANY_TO_VARIANT(in := #Setup, err => #temp16ReturnValue);
           // Validate Setup DB for the service control medium block and move to temp variable
           IF (#temp16ReturnValue = 0) THEN
               IF TypeOf(#tempVariant) = UDT_Service_ControlBlockMedium THEN
                   #temp16ReturnValue := MOVE_BLK_VARIANT(SRC := #tempVariant, COUNT := 1, SRC_INDEX := 0, DEST_INDEX := 0, DEST => #tempSetup);
               END_IF;
           END_IF;
       END_REGION

       REGION Configuration parameters
           //Initialize the used variable values
           #temp32TempDword1 := 16#1;
           #temp16IndexAnalog := 16#0;
           //#ConfigParaType.IndexAnalog := 16#0;
           #temp16IndexDigital := 16#0;
           //#ConfigParaType.IndexDigital := 16#0;
           #temp16IndexBinary := 16#0;
           //#ConfigParaType.IndexBinary := 16#0;
           #temp16IndexString := 16#0;
           //#ConfigParaType.IndexString := 16#0;
           //Used/Mapped parameter count with individual parameter type will written from the Tool
           #statTotalConfigParameters := #MAPPED_CONFIG_ANALOG + #MAPPED_CONFIG_DIGITAL + #MAPPED_CONFIG_BINARY + #MAPPED_CONFIG_STRING - 1;//Calculate the total used parameter
           IF ((#statTotalConfigParameters >= 0) AND (#statTotalConfigParameters <= #CONFIG_PARAMETER_MAX))  THEN
               FOR #temp16IndexOfDefinition := #CONFIG_PARAMETER_MIN TO #statTotalConfigParameters BY 1 DO//32 config parameters for Medium block.
                   #temp16ParameterCMAddress := BYTE_TO_INT(#tempSetup.configurationParameterData.definition[#temp16IndexOfDefinition].controlModule);//Get CM details from the setup DB.
                   #temp16ParameterType := #tempSetup.configurationParameterData.definition[#temp16IndexOfDefinition].type;//Get parameter type from the setup DB.
                   #temp16IndexMTP := #tempSetup.configurationParameterData.definition[#temp16IndexOfDefinition].indexMTP;//Get parameter indexMTP(wrapper DB) from the setup DB.
                   #temp16IndexIO := #tempSetup.configurationParameterData.definition[#temp16IndexOfDefinition].indexIO;//Get parameter indexIO(service block output config parameter) from the setup DB.
                   #tempUsed := #tempSetup.configurationParameterData.used;//Get parameter used info from setup DB
                   //Condition TO check CMs AND parameter types are in the range
                   IF (#temp16ParameterCMAddress <> 255) AND (#temp16ParameterCMAddress >= #NUMBER_OF_CONTROLMODULES_MIN) AND (#temp16ParameterCMAddress <= #NUMBER_OF_CONTROLMODULES)
                       AND (#temp16ParameterType >= #TYPE_NONE) AND (#temp16ParameterType <= #TYPE_STRING) THEN
                       #temp16TempInt1 := #temp16ParameterCMAddress / 32;    //DWORD - Adress
                       #temp16TempInt2 := #temp16ParameterCMAddress MOD 32;  //Bit - Adress
                       //If parameter is forced (FRC) --> Parameter is used
                       IF (((#tempUsed[#temp16TempInt1] AND SHL(IN := #temp32TempDword1, N := INT_TO_UINT(#temp16TempInt2))) <> 0) = TRUE) THEN
                           CASE #temp16ParameterType OF
                                   // If Parameter type = 1(Analog)
                               #TYPE_ANALOG:
                                   REGION Analog
                                       //Bit Masking funtionality for calculate the used Analog parameter
                                       #ConfigParaType.IndexAnalog := #ConfigParaType.IndexAnalog OR SHL(IN := #temp32TempDword1, N := INT_TO_UINT(#temp16IndexOfDefinition));
                                       //Condition to check the config analog parameters are within range 
                                       IF ((#temp16IndexIO >= #CONFIG_PARAMETER_MIN) AND (#temp16IndexIO <= #MAPPED_CONFIG_ANALOG)) THEN
                                           //WinCC Parameter View Faceplate logic
                                           #ConfigAna[#temp16IndexAnalog].WQC := #ConfigurationParameterAnalog[#temp16IndexMTP].WQC;
                                           #ConfigAna[#temp16IndexAnalog].ApplyEn := #ConfigurationParameterAnalog[#temp16IndexMTP].ApplyEn;
                                           #ConfigAna[#temp16IndexAnalog].ApplyInt := #ConfigurationParameterAnalog[#temp16IndexMTP].ApplyInt;
                                           #ConfigAna[#temp16IndexAnalog].StateChannel := #ConfigurationParameterAnalog[#temp16IndexMTP].StateChannel;
                                           #ConfigAna[#temp16IndexAnalog].StateOffAut := #ConfigurationParameterAnalog[#temp16IndexMTP].StateOffAut;
                                           #ConfigAna[#temp16IndexAnalog].StateOpAut := #ConfigurationParameterAnalog[#temp16IndexMTP].StateOpAut;
                                           #ConfigAna[#temp16IndexAnalog].StateAutAut := #ConfigurationParameterAnalog[#temp16IndexMTP].StateAutAut;
                                           #ConfigAna[#temp16IndexAnalog].StateOffAct := #ConfigurationParameterAnalog[#temp16IndexMTP].StateOffAct;
                                           #ConfigAna[#temp16IndexAnalog].StateOpAct := #ConfigurationParameterAnalog[#temp16IndexMTP].StateOpAct;
                                           #ConfigAna[#temp16IndexAnalog].StateAutAct := #ConfigurationParameterAnalog[#temp16IndexMTP].StateAutAct;
                                           #ConfigAna[#temp16IndexAnalog].SrcChannel := #ConfigurationParameterAnalog[#temp16IndexMTP].SrcChannel;
                                           #ConfigAna[#temp16IndexAnalog].SrcExtAut := #ConfigurationParameterAnalog[#temp16IndexMTP].SrcExtAut;
                                           #ConfigAna[#temp16IndexAnalog].SrcIntAut := #ConfigurationParameterAnalog[#temp16IndexMTP].SrcIntAut;
                                           #ConfigAna[#temp16IndexAnalog].SrcIntAct := #ConfigurationParameterAnalog[#temp16IndexMTP].SrcIntAct;
                                           #ConfigAna[#temp16IndexAnalog].SrcExtAct := #ConfigurationParameterAnalog[#temp16IndexMTP].SrcExtAct;
                                           #ConfigAna[#temp16IndexAnalog].VInt := #ConfigurationParameterAnalog[#temp16IndexMTP].VInt;
                                           #ConfigAna[#temp16IndexAnalog].VReq := #ConfigurationParameterAnalog[#temp16IndexMTP].VReq;
                                           #ConfigAna[#temp16IndexAnalog].VOut := #ConfigurationParameterAnalog[#temp16IndexMTP].VOut;
                                           #ConfigAna[#temp16IndexAnalog].VFbk := #ConfigurationParameterAnalog[#temp16IndexMTP].VFbk;
                                           #ConfigAna[#temp16IndexAnalog].VSclMin := #ConfigurationParameterAnalog[#temp16IndexMTP].VSclMin;
                                           #ConfigAna[#temp16IndexAnalog].VSclMax := #ConfigurationParameterAnalog[#temp16IndexMTP].VSclMax;
                                           #ConfigAna[#temp16IndexAnalog].VUnit := #ConfigurationParameterAnalog[#temp16IndexMTP].VUnit;
                                           #ConfigAna[#temp16IndexAnalog].VMin := #ConfigurationParameterAnalog[#temp16IndexMTP].VMin;
                                           #ConfigAna[#temp16IndexAnalog].VMax := #ConfigurationParameterAnalog[#temp16IndexMTP].VMax;
                                           //Write values from WinCC
                                           IF #ConfigurationParameterAnalog[#temp16IndexMTP].OSLevel = #StatConfigAnalog[#temp16IndexAnalog].OSLevel THEN
                                               #ConfigurationParameterAnalog[#temp16IndexMTP].OSLevel := #ConfigAna[#temp16IndexAnalog].OSLevel;
                                           ELSE
                                               #ConfigAna[#temp16IndexAnalog].OSLevel := #ConfigurationParameterAnalog[#temp16IndexMTP].OSLevel;
                                           END_IF;
                                           IF #ConfigurationParameterAnalog[#temp16IndexMTP].ApplyExt = #StatConfigAnalog[#temp16IndexAnalog].ApplyExt THEN
                                               #ConfigurationParameterAnalog[#temp16IndexMTP].ApplyExt := #ConfigAna[#temp16IndexAnalog].ApplyExt;
                                           ELSE
                                               #ConfigAna[#temp16IndexAnalog].ApplyExt := #ConfigurationParameterAnalog[#temp16IndexMTP].ApplyExt;
                                           END_IF;
                                           IF #ConfigurationParameterAnalog[#temp16IndexMTP].ApplyOp = #StatConfigAnalog[#temp16IndexAnalog].ApplyOp THEN
                                               #ConfigurationParameterAnalog[#temp16IndexMTP].ApplyOp := #ConfigAna[#temp16IndexAnalog].ApplyOp;
                                           ELSE
                                               #ConfigAna[#temp16IndexAnalog].ApplyOp := #ConfigurationParameterAnalog[#temp16IndexMTP].ApplyOp;
                                           END_IF;
                                           IF #ConfigurationParameterAnalog[#temp16IndexMTP].Sync = #StatConfigAnalog[#temp16IndexAnalog].Sync THEN
                                               #ConfigurationParameterAnalog[#temp16IndexMTP].Sync := #ConfigAna[#temp16IndexAnalog].Sync;
                                           ELSE
                                               #ConfigAna[#temp16IndexAnalog].Sync := #ConfigurationParameterAnalog[#temp16IndexMTP].Sync;
                                           END_IF;
                                           IF #ConfigurationParameterAnalog[#temp16IndexMTP].StateOffOp = #StatConfigAnalog[#temp16IndexAnalog].StateOffOp THEN
                                               #ConfigurationParameterAnalog[#temp16IndexMTP].StateOffOp := #ConfigAna[#temp16IndexAnalog].StateOffOp;
                                           ELSE
                                               #ConfigAna[#temp16IndexAnalog].StateOffOp := #ConfigurationParameterAnalog[#temp16IndexMTP].StateOffOp;
                                           END_IF;
                                           IF #ConfigurationParameterAnalog[#temp16IndexMTP].StateOpOp = #StatConfigAnalog[#temp16IndexAnalog].StateOpOp THEN
                                               #ConfigurationParameterAnalog[#temp16IndexMTP].StateOpOp := #ConfigAna[#temp16IndexAnalog].StateOpOp;
                                           ELSE
                                               #ConfigAna[#temp16IndexAnalog].StateOpOp := #ConfigurationParameterAnalog[#temp16IndexMTP].StateOpOp;
                                           END_IF;
                                           IF #ConfigurationParameterAnalog[#temp16IndexMTP].StateAutOp = #StatConfigAnalog[#temp16IndexAnalog].StateAutOp THEN
                                               #ConfigurationParameterAnalog[#temp16IndexMTP].StateAutOp := #ConfigAna[#temp16IndexAnalog].StateAutOp;
                                           ELSE
                                               #ConfigAna[#temp16IndexAnalog].StateAutOp := #ConfigurationParameterAnalog[#temp16IndexMTP].StateAutOp;
                                           END_IF;
                                           IF #ConfigurationParameterAnalog[#temp16IndexMTP].SrcIntOp = #StatConfigAnalog[#temp16IndexAnalog].SrcIntOp THEN
                                               #ConfigurationParameterAnalog[#temp16IndexMTP].SrcIntOp := #ConfigAna[#temp16IndexAnalog].SrcIntOp;
                                           ELSE
                                               #ConfigAna[#temp16IndexAnalog].SrcIntOp := #ConfigurationParameterAnalog[#temp16IndexMTP].SrcIntOp;
                                           END_IF;
                                           IF #ConfigurationParameterAnalog[#temp16IndexMTP].SrcExtOp = #StatConfigAnalog[#temp16IndexAnalog].SrcExtOp THEN
                                               #ConfigurationParameterAnalog[#temp16IndexMTP].SrcExtOp := #ConfigAna[#temp16IndexAnalog].SrcExtOp;
                                           ELSE
                                               #ConfigAna[#temp16IndexAnalog].SrcExtOp := #ConfigurationParameterAnalog[#temp16IndexMTP].SrcExtOp;
                                           END_IF;
                                           IF #ConfigurationParameterAnalog[#temp16IndexMTP].VExt = #StatConfigAnalog[#temp16IndexAnalog].VExt THEN
                                               #ConfigurationParameterAnalog[#temp16IndexMTP].VExt := #ConfigAna[#temp16IndexAnalog].VExt;
                                           ELSE
                                               #ConfigAna[#temp16IndexAnalog].VExt := #ConfigurationParameterAnalog[#temp16IndexMTP].VExt;
                                           END_IF;
                                           IF #ConfigurationParameterAnalog[#temp16IndexMTP].VOp = #StatConfigAnalog[#temp16IndexAnalog].VOp THEN
                                               #ConfigurationParameterAnalog[#temp16IndexMTP].VOp := #ConfigAna[#temp16IndexAnalog].VOp;
                                           ELSE
                                               #ConfigAna[#temp16IndexAnalog].VOp := #ConfigurationParameterAnalog[#temp16IndexMTP].VOp;
                                           END_IF;

                                           #StatConfigAnalog[#temp16IndexAnalog].OSLevel := #ConfigAna[#temp16IndexAnalog].OSLevel;
                                           #StatConfigAnalog[#temp16IndexAnalog].ApplyExt := #ConfigAna[#temp16IndexAnalog].ApplyExt;
                                           #StatConfigAnalog[#temp16IndexAnalog].ApplyOp := #ConfigAna[#temp16IndexAnalog].ApplyOp;
                                           #StatConfigAnalog[#temp16IndexAnalog].Sync := #ConfigAna[#temp16IndexAnalog].Sync;
                                           #StatConfigAnalog[#temp16IndexAnalog].StateOffOp := #ConfigAna[#temp16IndexAnalog].StateOffOp;
                                           #StatConfigAnalog[#temp16IndexAnalog].StateOpOp := #ConfigAna[#temp16IndexAnalog].StateOpOp;
                                           #StatConfigAnalog[#temp16IndexAnalog].StateAutOp := #ConfigAna[#temp16IndexAnalog].StateAutOp;
                                           #StatConfigAnalog[#temp16IndexAnalog].SrcIntOp := #ConfigAna[#temp16IndexAnalog].SrcIntOp;
                                           #StatConfigAnalog[#temp16IndexAnalog].SrcExtOp := #ConfigAna[#temp16IndexAnalog].SrcExtOp;
                                           #StatConfigAnalog[#temp16IndexAnalog].VExt := #ConfigAna[#temp16IndexAnalog].VExt;
                                           #StatConfigAnalog[#temp16IndexAnalog].VOp := #ConfigAna[#temp16IndexAnalog].VOp;
                                       END_IF;
                                       #temp16IndexAnalog := #temp16IndexAnalog + 1;
                                   END_REGION
                                   // If Parameter type = 2(Digital)
                               #TYPE_DIGITAL:
                                   REGION Digital
                                       //Bit Masking funtionality for calculate the used Digital parameter
                                       #ConfigParaType.IndexDigital := #ConfigParaType.IndexDigital OR SHL(IN := #temp32TempDword1, N := INT_TO_UINT(#temp16IndexOfDefinition));
                                       //Condition to check the config digital parameters are within range 
                                       IF ((#temp16IndexIO >= #CONFIG_PARAMETER_MIN) AND (#temp16IndexIO <= #MAPPED_CONFIG_DIGITAL)) THEN
                                           //WinCC Parameter View Faceplate logic
                                           #ConfigDint[#temp16IndexDigital].WQC := #ConfigurationParameterDigital[#temp16IndexMTP].WQC;
                                           #ConfigDint[#temp16IndexDigital].ApplyEn := #ConfigurationParameterDigital[#temp16IndexMTP].ApplyEn;
                                           #ConfigDint[#temp16IndexDigital].ApplyInt := #ConfigurationParameterDigital[#temp16IndexMTP].ApplyInt;
                                           #ConfigDint[#temp16IndexDigital].StateChannel := #ConfigurationParameterDigital[#temp16IndexMTP].StateChannel;
                                           #ConfigDint[#temp16IndexDigital].StateOffAut := #ConfigurationParameterDigital[#temp16IndexMTP].StateOffAut;
                                           #ConfigDint[#temp16IndexDigital].StateOpAut := #ConfigurationParameterDigital[#temp16IndexMTP].StateOpAut;
                                           #ConfigDint[#temp16IndexDigital].StateAutAut := #ConfigurationParameterDigital[#temp16IndexMTP].StateAutAut;
                                           #ConfigDint[#temp16IndexDigital].StateOffAct := #ConfigurationParameterDigital[#temp16IndexMTP].StateOffAct;
                                           #ConfigDint[#temp16IndexDigital].StateOpAct := #ConfigurationParameterDigital[#temp16IndexMTP].StateOpAct;
                                           #ConfigDint[#temp16IndexDigital].StateAutAct := #ConfigurationParameterDigital[#temp16IndexMTP].StateAutAct;
                                           #ConfigDint[#temp16IndexDigital].SrcChannel := #ConfigurationParameterDigital[#temp16IndexMTP].SrcChannel;
                                           #ConfigDint[#temp16IndexDigital].SrcExtAut := #ConfigurationParameterDigital[#temp16IndexMTP].SrcExtAut;
                                           #ConfigDint[#temp16IndexDigital].SrcIntAut := #ConfigurationParameterDigital[#temp16IndexMTP].SrcIntAut;
                                           #ConfigDint[#temp16IndexDigital].SrcIntAct := #ConfigurationParameterDigital[#temp16IndexMTP].SrcIntAct;
                                           #ConfigDint[#temp16IndexDigital].SrcExtAct := #ConfigurationParameterDigital[#temp16IndexMTP].SrcExtAct;
                                           #ConfigDint[#temp16IndexDigital].VInt := #ConfigurationParameterDigital[#temp16IndexMTP].VInt;
                                           #ConfigDint[#temp16IndexDigital].VReq := #ConfigurationParameterDigital[#temp16IndexMTP].VReq;
                                           #ConfigDint[#temp16IndexDigital].VOut := #ConfigurationParameterDigital[#temp16IndexMTP].VOut;
                                           #ConfigDint[#temp16IndexDigital].VFbk := #ConfigurationParameterDigital[#temp16IndexMTP].VFbk;
                                           #ConfigDint[#temp16IndexDigital].VSclMin := #ConfigurationParameterDigital[#temp16IndexMTP].VSclMin;
                                           #ConfigDint[#temp16IndexDigital].VSclMax := #ConfigurationParameterDigital[#temp16IndexMTP].VSclMax;
                                           #ConfigDint[#temp16IndexDigital].VUnit := #ConfigurationParameterDigital[#temp16IndexMTP].VUnit;
                                           #ConfigDint[#temp16IndexDigital].VMin := #ConfigurationParameterDigital[#temp16IndexMTP].VMin;
                                           #ConfigDint[#temp16IndexDigital].VMax := #ConfigurationParameterDigital[#temp16IndexMTP].VMax;
                                           //Write values from WinCC
                                           IF #ConfigurationParameterDigital[#temp16IndexMTP].OSLevel = #StatConfigDigital[#temp16IndexDigital].OSLevel THEN
                                               #ConfigurationParameterDigital[#temp16IndexMTP].OSLevel := #ConfigDint[#temp16IndexDigital].OSLevel;
                                           ELSE
                                               #ConfigDint[#temp16IndexDigital].OSLevel := #ConfigurationParameterDigital[#temp16IndexMTP].OSLevel;
                                           END_IF;
                                           IF #ConfigurationParameterDigital[#temp16IndexMTP].ApplyExt = #StatConfigDigital[#temp16IndexDigital].ApplyExt THEN
                                               #ConfigurationParameterDigital[#temp16IndexMTP].ApplyExt := #ConfigDint[#temp16IndexDigital].ApplyExt;
                                           ELSE
                                               #ConfigDint[#temp16IndexDigital].ApplyExt := #ConfigurationParameterDigital[#temp16IndexMTP].ApplyExt;
                                           END_IF;
                                           IF #ConfigurationParameterDigital[#temp16IndexMTP].ApplyOp = #StatConfigDigital[#temp16IndexDigital].ApplyOp THEN
                                               #ConfigurationParameterDigital[#temp16IndexMTP].ApplyOp := #ConfigDint[#temp16IndexDigital].ApplyOp;
                                           ELSE
                                               #ConfigDint[#temp16IndexDigital].ApplyOp := #ConfigurationParameterDigital[#temp16IndexMTP].ApplyOp;
                                           END_IF;
                                           IF #ConfigurationParameterDigital[#temp16IndexMTP].Sync = #StatConfigDigital[#temp16IndexDigital].Sync THEN
                                               #ConfigurationParameterDigital[#temp16IndexMTP].Sync := #ConfigDint[#temp16IndexDigital].Sync;
                                           ELSE
                                               #ConfigDint[#temp16IndexDigital].Sync := #ConfigurationParameterDigital[#temp16IndexMTP].Sync;
                                           END_IF;
                                           IF #ConfigurationParameterDigital[#temp16IndexMTP].StateOffOp = #StatConfigDigital[#temp16IndexDigital].StateOffOp THEN
                                               #ConfigurationParameterDigital[#temp16IndexMTP].StateOffOp := #ConfigDint[#temp16IndexDigital].StateOffOp;
                                           ELSE
                                               #ConfigDint[#temp16IndexDigital].StateOffOp := #ConfigurationParameterDigital[#temp16IndexMTP].StateOffOp;
                                           END_IF;
                                           IF #ConfigurationParameterDigital[#temp16IndexMTP].StateOpOp = #StatConfigDigital[#temp16IndexDigital].StateOpOp THEN
                                               #ConfigurationParameterDigital[#temp16IndexMTP].StateOpOp := #ConfigDint[#temp16IndexDigital].StateOpOp;
                                           ELSE
                                               #ConfigDint[#temp16IndexDigital].StateOpOp := #ConfigurationParameterDigital[#temp16IndexMTP].StateOpOp;
                                           END_IF;
                                           IF #ConfigurationParameterDigital[#temp16IndexMTP].StateAutOp = #StatConfigDigital[#temp16IndexDigital].StateAutOp THEN
                                               #ConfigurationParameterDigital[#temp16IndexMTP].StateAutOp := #ConfigDint[#temp16IndexDigital].StateAutOp;
                                           ELSE
                                               #ConfigDint[#temp16IndexDigital].StateAutOp := #ConfigurationParameterDigital[#temp16IndexMTP].StateAutOp;
                                           END_IF;
                                           IF #ConfigurationParameterDigital[#temp16IndexMTP].SrcIntOp = #StatConfigDigital[#temp16IndexDigital].SrcIntOp THEN
                                               #ConfigurationParameterDigital[#temp16IndexMTP].SrcIntOp := #ConfigDint[#temp16IndexDigital].SrcIntOp;
                                           ELSE
                                               #ConfigDint[#temp16IndexDigital].SrcIntOp := #ConfigurationParameterDigital[#temp16IndexMTP].SrcIntOp;
                                           END_IF;
                                           IF #ConfigurationParameterDigital[#temp16IndexMTP].SrcExtOp = #StatConfigDigital[#temp16IndexDigital].SrcExtOp THEN
                                               #ConfigurationParameterDigital[#temp16IndexMTP].SrcExtOp := #ConfigDint[#temp16IndexDigital].SrcExtOp;
                                           ELSE
                                               #ConfigDint[#temp16IndexDigital].SrcExtOp := #ConfigurationParameterDigital[#temp16IndexMTP].SrcExtOp;
                                           END_IF;
                                           IF #ConfigurationParameterDigital[#temp16IndexMTP].VExt = #StatConfigDigital[#temp16IndexDigital].VExt THEN
                                               #ConfigurationParameterDigital[#temp16IndexMTP].VExt := #ConfigDint[#temp16IndexDigital].VExt;
                                           ELSE
                                               #ConfigDint[#temp16IndexDigital].VExt := #ConfigurationParameterDigital[#temp16IndexMTP].VExt;
                                           END_IF;
                                           IF #ConfigurationParameterDigital[#temp16IndexMTP].VOp = #StatConfigDigital[#temp16IndexDigital].VOp THEN
                                               #ConfigurationParameterDigital[#temp16IndexMTP].VOp := #ConfigDint[#temp16IndexDigital].VOp;
                                           ELSE
                                               #ConfigDint[#temp16IndexDigital].VOp := #ConfigurationParameterDigital[#temp16IndexMTP].VOp;
                                           END_IF;

